// TIA Portal project "Project112" (V16)

(* hardware
DEVICE "S71500/ET200MP station_1"  S7-1500 station
   slot 0: "Rail_0"  Rack  6ES7 590-1***0-0AA0
   slot 0: "PS 25W 24VDC_1"  PS 25W 24VDC  6ES7 505-0KA00-0AB0  V1.0
   slot 1: "fillingStation"  CPU 1511F-1 PN  6ES7 511-1FK00-0AB0  V1.8
      slot 3: "CPU display_1"  6ES7591-1AA00-0AA0
      slot 32768: "PROFINET interface_1"  X1
         slot 32769: "Port_1"  X1 P1
         slot 32770: "Port_2"  X1 P2
   slot 2: "DI 16x24VDC BA_1"  DI 16x24VDC BA  6ES7 521-1BH10-0AA0  V1.1
   slot 3: "DQ 8x24VDC/2A HF_1"  DQ 8x24VDC/2A HF  6ES7 522-1BF00-0AB0  V2.2
   slot 4: "AI 4xU/I/RTD/TC ST_1"  AI 4xU/I/RTD/TC ST  6ES7 531-7QD00-0AB0  V1.0
DEVICE "HMI_1"  TP700 Comfort
   slot 0: "HMI_1"  TP700 Comfort  6AV2 124-0GC01-0AX0  16.0.0.0
   slot 1: "HMI_RT_1"  TP700 Comfort  6AV2 124-0GC01-0AX0  16.0.0.0
   slot 5: "HMI_1.IE_CP_1"  PROFINET Interface  16.0.0.0
      slot 1: "PROFINET Interface_1"  PROFINET Interface
         slot 1: "Port_1"  Port
         slot 2: "Port_2"  Port
   slot 7: "HMI_1.MPI/DP_CP_1"  MPI/DP Interface  16.0.0.0
DEVICE "GSD device_1"  GSD.Device.PN
   slot 0: "Rack"  Rack  V1.0
   slot 0: "SINAMICS-G120-CU240E-2PN"  SINAMICS G120 CU240E-2 PN(-F) V4.5  6SL3 244-0BB1x-1FAx  V4.5
      slot 0: "SINAMICS G120 CU240E-2 PN(-F) V4.5"  SINAMICS G120 CU240E-2 PN(-F) V4.5
      slot 1: "PN-IO"  PN-IO
         slot 1: "Port 1"  Port 1
         slot 2: "Port 2"  Port 2
      slot 1: "Drive_1"  Drive
         slot 0: "Module Access Point"  Module Access Point
   slot 2: "Free telegram, PZD-8/8"  Free telegram, PZD-8/8
*)

// ===== PLC "fillingStation"  CPU 1511F-1 PN =====

VAR_GLOBAL   // PLC tag table "Default tag table"
   "Emg_stop" AT %I0.0 : Bool;
   "Start" AT %I0.1 : Bool;
   "b01_highlevel" AT %I0.2 : Bool;
   "bo2_lowlevel" AT %I0.3 : Bool;
   "pompe_km1" AT %Q0.0 : Bool;
   "valvefilling_1" AT %Q0.1 : Bool;
   "valvefilling_2" AT %Q0.2 : Bool;
   "evacuation_valve" AT %Q0.3 : Bool;
   "stop_bt" AT %M0.0 : Bool;
   "stop_bt(1)" AT %M0.7 : Bool;
   "statehandler" AT %M0.1 : Bool;
   "generalErrors" AT %MD10 : DWord;
   "pompeerror" AT %M10.0 : Bool;
   "pompe_error" AT %M0.2 : Bool;
   "System_Byte" AT %MB1 : Byte;
   "FirstScan" AT %M1.0 : Bool;
   "DiagStatusUpdate" AT %M1.1 : Bool;
   "AlwaysTRUE" AT %M1.2 : Bool;
   "AlwaysFALSE" AT %M1.3 : Bool;
   "System_Byte(1)" AT %MB1 : Byte;
   "Clock_Byte" AT %MB0 : Byte;
   "Clock_10Hz" AT %M0.0 : Bool;
   "Clock_5Hz" AT %M0.1 : Bool;
   "Clock_2.5Hz" AT %M0.2 : Bool;
   "Clock_2Hz" AT %M0.3 : Bool;
   "Clock_1.25Hz" AT %M0.4 : Bool;
   "Clock_1Hz" AT %M0.5 : Bool;
   "Clock_0.625Hz" AT %M0.6 : Bool;
   "Clock_0.5Hz" AT %M0.7 : Bool;
   "actual_wight_card" AT %IW2 : Int;
END_VAR

VAR_GLOBAL   // PLC tag table "input"
   "start(1)" AT %I0.4 : Bool;
   "stop" AT %I0.5 : Bool;
   "reset" AT %I0.6 : Bool;
   "box_detection" AT %I0.7 : Bool;
   "box_at_filling" AT %I1.0 : Bool;
   "box_at_scale" AT %I1.1 : Bool;
   "box_reject" AT %I1.2 : Bool;
   "box_left" AT %I1.3 : Bool;
   "reject_cyl_extended" AT %I1.4 : Bool;
   "reject_cyl_retracted" AT %I1.5 : Bool;
   "caping_cylinder_extended" AT %I1.6 : Bool;
   "caping_cylinder_retracted" AT %I1.7 : Bool;
   "inspect_ol" AT %I2.0 : Bool;
   "conveyer_moving" AT %I2.1 : Bool;
   "valve_switch_open" AT %I2.2 : Bool;
   "main_air_switch" AT %I2.7 : Bool;
   "main_valve_open_fb" AT %I3.1 : Bool;
   "input_vfd" AT %I500.0 : "udt_vfd_status";
   "filling_cyl_retracted" AT %I4.0 : Bool;
   "filling_cyl_extended" AT %I4.1 : Bool;
   "curent_speed" AT %IW600 : Word;
   "part_at_sealing" AT %I3.2 : Bool;
   "cap_carrier_extended" AT %I4.2 : Bool;
   "cap_carrier_retracted" AT %I4.3 : Bool;
   "filling_valve_extended" AT %I4.4 : Bool;
   "filling_valve_retracted" AT %I4.5 : Bool;
   "sealing_locater_extended" AT %I4.6 : Bool;
   "sealing_locater_retacted" AT %I4.7 : Bool;
   "cap_valve_open" AT %I5.0 : Bool;
   "box_at_reject" AT %I5.1 : Bool;
END_VAR

VAR_GLOBAL   // PLC tag table "output"
   "Ev_valve_refill" AT %Q1.0 : Bool;
   "EV_capping" AT %Q1.1 : Bool;
   "EV_capping_return" AT %Q1.2 : Bool;
   "Ev_reject_cylinder" AT %Q1.3 : Bool;
   "main_air_valve" AT %Q1.4 : Bool;
   "tower_green" AT %Q1.5 : Bool;
   "tower_red" AT %Q1.6 : Bool;
   "tower_orange" AT %Q1.7 : Bool;
   "tower_buzer" AT %Q2.0 : Bool;
   "udt_vfd_cmd" AT %Q500.0 : "vfd_cmd";
   "ev_filling_cylinder" AT %Q2.1 : Bool;
   "set_point_vfd" AT %QW600 : Word;
   "cap_motor" AT %Q2.2 : Bool;
   "ev_filling_valve_cyl" AT %Q2.3 : Bool;
   "ev_cap_valve_carrier_cyl" AT %Q2.4 : Bool;
END_VAR

TYPE "udt_state_handler"
   STRUCT
      status : Struct
         ready : Bool;
         running : Bool;
         faulted : Bool;
         stop : Bool;
         safety_ok : Bool;
         air_ok : Bool;
      END_STRUCT;
      cmd : Struct
         reset : Bool;
         start : Bool;
         stop : Bool;
      END_STRUCT;
      cnf : Struct
         state : Int;
      END_STRUCT;
      flts : Struct
         air_system_faulted : Bool;
         safety_emg_stop_btn : Bool;
      END_STRUCT;
   END_STRUCT;
END_TYPE

TYPE "udt_tower_handler"
   STRUCT
      status : Struct
         running : Bool;
         faulted : Bool;
         stop : Bool;
      END_STRUCT;
      cmd : Struct
         turn_red : Bool;
         turn_green : Bool;
         turn_orange : Bool;
         turn_bazer : Bool;
      END_STRUCT;
      flt : Struct
         x_sparte : Bool;
      END_STRUCT;
      cnf : Struct
         x_spare : Bool;
      END_STRUCT;
   END_STRUCT;
END_TYPE

TYPE "udt_equipement"
   STRUCT
      state : Struct
         running : Bool;
         reject_done : Bool;
         filling_done : Bool;
         sealing_done : Bool;
         varification_done : Bool;
         faulted : Bool;
         ready : Bool;
         part_detected : Bool;
         state : Int;
      END_STRUCT;
      cmd : Struct
         converyer_cmd : Bool;
         "filling _valve_cmd" : Bool;
         cmd_cylinder_filling : Bool;
         cmd_cylinder_sealing : Bool;
         cmd_sealing_motor : Bool;
         cmd_cylinder_reject : Bool;
         cmd_trigger_verificaiton : Bool;
         enable_filling : Bool;
         enable_sealing : Bool;
         enable_verification : Bool;
         enable_reject : Bool;
      END_STRUCT;
      flt : Struct
         main_sequece_timeout : Bool;
      END_STRUCT;
      cnf : Struct
         scale_pass_weight : Int := 200;
      END_STRUCT;
   END_STRUCT;
END_TYPE

TYPE "filling_station_udt"
   STRUCT
      status : Struct
         cyl_at_retract : Bool;
         cyl_at_extened : Bool;
         part_at_felling : Bool;
         running : Bool;
         faulted : Bool;
         felling_done : Bool;
         felling_start : Bool;
         valve_open : Bool;
         cyl_valve_at_retract : Bool;
         cyl_valve_at_extend : Bool;
         state : Int;
      END_STRUCT;
      cmd : Struct
         locater_cylinder_cmd : Bool;
         valve_open_cmd : Bool;
         valve_cylinder_cmd : Bool;
      END_STRUCT;
      flt_valve : Word;   // these will define the faults of the valve
      flt2 : Word;   // these are for the filling valve carrier cylinder
      flt1 : Word;   // these are for filling locater cylinder
      cfg : Struct
         valve_open_time : Time := T#10ms;
      END_STRUCT;
   END_STRUCT;
END_TYPE

TYPE "sealing_udt"
   STRUCT
      status : Struct
         cap_carrier_retract : Bool;
         cap_carrier_extended : Bool;
         cyl_at_retract : Bool;
         cyl_at_extended : Bool;
         running : Bool;
         stoped : Bool;
         part_at_sealing : Bool;
         motor_running : Bool;
         cap_present : Bool;
         state : Int;
         open_cap_valve : Int;
      END_STRUCT;
      cmd : Struct
         motor_start_cmd : Bool;
         locater_cyl_cmd : Bool;
         cap_carring_cyl_cmd : Bool;
         open_cap_valve_cmd : Bool;
      END_STRUCT;
      flt_valve : Word;
      flt_valve_carrier_cyl : Word;
      flt_locater_cylinder : Word;
      cnf : Struct
         spare : Bool;
      END_STRUCT;
   END_STRUCT;
END_TYPE

TYPE "scaling_udt"
   STRUCT
      status : Struct
         actual_weight_bottle : Int;
         running : Bool;
         stop : Bool;
         pass_part : Bool;
         reject_part : Bool;
      END_STRUCT;
      cmd : Struct
         spare : Bool;
      END_STRUCT;
      cnf : Struct
         max_weight : Int := 140;
         min_weight : Int := 150;
      END_STRUCT;
      flt : Word;
   END_STRUCT;
END_TYPE

TYPE "reject_udt"
   STRUCT
      status : Struct
         cyl_at_retract : Bool;
         cyl_at_extend : Bool;
         running : Bool;
         faulted : Bool;
         state : Int;
      END_STRUCT;
      cmd : Struct
         spare : Bool;
      END_STRUCT;
      flt : Word;
      cnf : Struct
         reject_count : Int;
      END_STRUCT;
   END_STRUCT;
END_TYPE

TYPE "udt_vfd_status"
   STRUCT
      "Ready to switch on" : Bool;
      "Ready for operation" : Bool;
      "Operation enabled" : Bool;
      "Fault active" : Bool;
      "OFF2 inactive" : Bool;
      "OFF3 inactive" : Bool;
      "Switching-on inhibited" : Bool;
      "Warning active" : Bool;
      "Speed setpoint/actual value comparison" : Bool;
      "Control requested" : Bool;
      "Setpoint reached" : Bool;
      "Torque limit active" : Bool;
   END_STRUCT;
END_TYPE

TYPE "vfd_cmd"
   STRUCT
      "ON/OFF1" : Bool;
      OFF2 : Bool;
      OFF3 : Bool;
      "Enable operation" : Bool;
      "Enable ramp-function generator" : Bool;
      "Continue ramp-function generator" : Bool;
      "Enable setpoint" : Bool;
      "Acknowledge fault" : Bool;
      "Control by PLC" : Bool;
   END_STRUCT;
END_TYPE

TYPE "hmi_cmd_state"
   STRUCT
      cmd : Struct
         oprator_speed_setpoint : Int;
      END_STRUCT;
      status : Struct
         set_point_valid : Bool;
      END_STRUCT;
   END_STRUCT;
END_TYPE

DATA_BLOCK "Main_Safety_RTG1_DB"   // DB1, F_DB
{ S7_Optimized_Access := 'TRUE' }
NAME : FUSI
VERSION : 0.1
// stored: InstanceOfName Main_Safety_RTG1
"Main_Safety_RTG1"
BEGIN
END_DATA_BLOCK

DATA_BLOCK "global_data_block"   // DB6
{ S7_Optimized_Access := 'TRUE' }
VERSION : 0.1
   VAR
      verification_handler : "scaling_udt";
      reject_handler : "reject_udt";
      hmi_cmd_state : "hmi_cmd_state";
      sealing_handler : "sealing_udt";
      equipement_handler : "udt_equipement";
      filling_station_handler : "filling_station_udt";
      tower_handling : "udt_tower_handler";
      machine_state : "udt_state_handler";
   END_VAR
BEGIN
END_DATA_BLOCK

// folder: System blocks/Program resources

DATA_BLOCK "air_check"   // DB2
{ S7_Optimized_Access := 'TRUE' }
AUTHOR : Simatic
FAMILY : IEC
NAME : IEC_TMR
VERSION : 1.0
// stored: InstanceOfName IEC_TIMER
"IEC_TIMER"
BEGIN
END_DATA_BLOCK

DATA_BLOCK "verify_air_present"   // DB5
{ S7_Optimized_Access := 'TRUE' }
AUTHOR : Simatic
FAMILY : IEC
NAME : IEC_TMR
VERSION : 1.0
// stored: InstanceOfName IEC_TIMER
"IEC_TIMER"
BEGIN
END_DATA_BLOCK

DATA_BLOCK "valve_timing"   // DB15
{ S7_Optimized_Access := 'TRUE' }
AUTHOR : Simatic
FAMILY : IEC
NAME : IEC_TMR
VERSION : 1.0
// stored: InstanceOfName IEC_TIMER
"IEC_TIMER"
BEGIN
END_DATA_BLOCK

DATA_BLOCK "IEC_Timer_0_DB_1"   // DB16
{ S7_Optimized_Access := 'TRUE' }
AUTHOR : Simatic
FAMILY : IEC
NAME : IEC_TMR
VERSION : 1.0
// stored: InstanceOfName IEC_TIMER
"IEC_TIMER"
BEGIN
END_DATA_BLOCK

DATA_BLOCK "motor_time"   // DB17
{ S7_Optimized_Access := 'TRUE' }
AUTHOR : Simatic
FAMILY : IEC
NAME : IEC_TMR
VERSION : 1.0
// stored: InstanceOfName IEC_TIMER
"IEC_TIMER"
BEGIN
END_DATA_BLOCK

DATA_BLOCK "IEC_Timer_0_DB_2"   // DB18
{ S7_Optimized_Access := 'TRUE' }
AUTHOR : Simatic
FAMILY : IEC
NAME : IEC_TMR
VERSION : 1.0
// stored: InstanceOfName IEC_TIMER
"IEC_TIMER"
BEGIN
END_DATA_BLOCK

DATA_BLOCK "IEC_Timer_0_DB_3"   // DB19
{ S7_Optimized_Access := 'TRUE' }
AUTHOR : Simatic
FAMILY : IEC
NAME : IEC_TMR
VERSION : 1.0
// stored: InstanceOfName IEC_TIMER
"IEC_TIMER"
BEGIN
END_DATA_BLOCK

DATA_BLOCK "wire_break"   // DB20
{ S7_Optimized_Access := 'TRUE' }
AUTHOR : Simatic
FAMILY : IEC
NAME : IEC_TMR
VERSION : 1.0
// stored: InstanceOfName IEC_TIMER
"IEC_TIMER"
BEGIN
END_DATA_BLOCK

DATA_BLOCK "IEC_Timer_0_DB_4"   // DB21
{ S7_Optimized_Access := 'TRUE' }
AUTHOR : Simatic
FAMILY : IEC
NAME : IEC_TMR
VERSION : 1.0
// stored: InstanceOfName IEC_TIMER
"IEC_TIMER"
BEGIN
END_DATA_BLOCK

DATA_BLOCK "IEC_Timer_0_DB_5"   // DB22
{ S7_Optimized_Access := 'TRUE' }
AUTHOR : Simatic
FAMILY : IEC
NAME : IEC_TMR
VERSION : 1.0
// stored: InstanceOfName IEC_TIMER
"IEC_TIMER"
BEGIN
END_DATA_BLOCK

DATA_BLOCK "timeout]"   // DB25
{ S7_Optimized_Access := 'TRUE' }
AUTHOR : Simatic
FAMILY : IEC
NAME : IEC_TMR
VERSION : 1.0
// stored: InstanceOfName IEC_TIMER
"IEC_TIMER"
BEGIN
END_DATA_BLOCK

DATA_BLOCK "IEC_Timer_0_DB_8"   // DB26
{ S7_Optimized_Access := 'TRUE' }
AUTHOR : Simatic
FAMILY : IEC
NAME : IEC_TMR
VERSION : 1.0
// stored: InstanceOfName IEC_TIMER
"IEC_TIMER"
BEGIN
END_DATA_BLOCK

DATA_BLOCK "signal_che k"   // DB27
{ S7_Optimized_Access := 'TRUE' }
AUTHOR : Simatic
FAMILY : IEC
NAME : IEC_TMR
VERSION : 1.0
// stored: InstanceOfName IEC_TIMER
"IEC_TIMER"
BEGIN
END_DATA_BLOCK

DATA_BLOCK "cyl_extended_check"   // DB28
{ S7_Optimized_Access := 'TRUE' }
AUTHOR : Simatic
FAMILY : IEC
NAME : IEC_TMR
VERSION : 1.0
// stored: InstanceOfName IEC_TIMER
"IEC_TIMER"
BEGIN
END_DATA_BLOCK

DATA_BLOCK "cylinder"   // DB29
{ S7_Optimized_Access := 'TRUE' }
AUTHOR : Simatic
FAMILY : IEC
NAME : IEC_TMR
VERSION : 1.0
// stored: InstanceOfName IEC_TIMER
"IEC_TIMER"
BEGIN
END_DATA_BLOCK

DATA_BLOCK "IEC_Timer_0_DB_9"   // DB30
{ S7_Optimized_Access := 'TRUE' }
AUTHOR : Simatic
FAMILY : IEC
NAME : IEC_TMR
VERSION : 1.0
// stored: InstanceOfName IEC_TIMER
"IEC_TIMER"
BEGIN
END_DATA_BLOCK

DATA_BLOCK "setpoint"   // DB31
{ S7_Optimized_Access := 'TRUE' }
AUTHOR : Simatic
FAMILY : IEC
NAME : IEC_TMR
VERSION : 1.0
// stored: InstanceOfName IEC_TIMER
"IEC_TIMER"
BEGIN
END_DATA_BLOCK

DATA_BLOCK "IEC_Timer_0_DB_10"   // DB33
{ S7_Optimized_Access := 'TRUE' }
AUTHOR : Simatic
FAMILY : IEC
NAME : IEC_TMR
VERSION : 1.0
// stored: InstanceOfName IEC_TIMER
"IEC_TIMER"
BEGIN
END_DATA_BLOCK

// folder: equipement

DATA_BLOCK "filling_sequence_DB"   // DB11
{ S7_Optimized_Access := 'TRUE' }
VERSION : 0.1
// stored: InstanceOfName filling_sequence
"filling_sequence"
BEGIN
END_DATA_BLOCK

DATA_BLOCK "sealing_db"   // DB12
{ S7_Optimized_Access := 'TRUE' }
VERSION : 0.1
// stored: InstanceOfName sealing_sequnce
"sealing_sequnce"
BEGIN
END_DATA_BLOCK

DATA_BLOCK "scaling_sequence_DB"   // DB13
{ S7_Optimized_Access := 'TRUE' }
VERSION : 0.1
// stored: InstanceOfName scaling_sequence
"scaling_sequence"
BEGIN
END_DATA_BLOCK

DATA_BLOCK "1_main_squence_DB"   // DB32
{ S7_Optimized_Access := 'TRUE' }
VERSION : 0.1
// stored: InstanceOfName 1_main_squence
"1_main_squence"
BEGIN
END_DATA_BLOCK

// folder: machine

DATA_BLOCK "safety_block_DB"   // DB7
{ S7_Optimized_Access := 'TRUE' }
VERSION : 0.1
// stored: InstanceOfName safety_block
"safety_block"
BEGIN
END_DATA_BLOCK

DATA_BLOCK "air_management_blk_DB"   // DB8
{ S7_Optimized_Access := 'TRUE' }
VERSION : 0.1
// stored: InstanceOfName air_management_blk
"air_management_blk"
BEGIN
END_DATA_BLOCK

DATA_BLOCK "tower_handler_DB"   // DB9
{ S7_Optimized_Access := 'TRUE' }
VERSION : 0.1
// stored: InstanceOfName tower_handler
"tower_handler"
BEGIN
END_DATA_BLOCK

DATA_BLOCK "state_handler_DB"   // DB10
{ S7_Optimized_Access := 'TRUE' }
VERSION : 0.1
// stored: InstanceOfName state_handler
"state_handler"
BEGIN
END_DATA_BLOCK

// folder: (top level)

FUNCTION_BLOCK "Main_Safety_RTG1"   // FB1, F_FBD
{ S7_Optimized_Access := 'TRUE' }
BEGIN

REGION Network 1
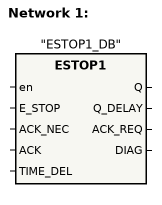
   "ESTOP1_DB"();   // ESTOP1
END_REGION
END_FUNCTION_BLOCK

ORGANIZATION_BLOCK "Main"   // OB1, LAD, ProgramCycle
TITLE = "Main Program Sweep (Cycle)"
{ S7_Optimized_Access := 'TRUE' }
VERSION : 0.1
   VAR_INPUT
      Initial_Call : Bool;   // Initial call of this OB
      Remanence : Bool;   // =True, if remanent data are available
   END_VAR
BEGIN

REGION Network 1: this the systeme process
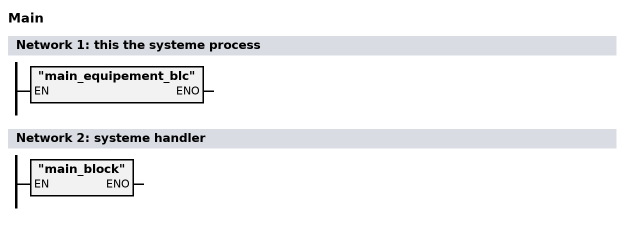
   RUNG wire#powerrail
      "main_equipement_blc"()
   END_RUNG
   // the same network as SCL:
   "main_equipement_blc"();
END_REGION

REGION Network 2: systeme handler
   RUNG wire#powerrail
      "main_block"()
   END_RUNG
   // the same network as SCL:
   "main_block"();
END_REGION

REGION Network 3: error handler block
END_REGION
END_ORGANIZATION_BLOCK

// folder: equipement

FUNCTION_BLOCK "1_main_squence"   // FB6, LAD
{ S7_Optimized_Access := 'TRUE' }
VERSION : 0.1
   VAR_INPUT
      conveyor_feedbak : Bool;
      part_at_filling : Bool;
      part_at_sealing : Bool;
      part_verification : Bool;
      part_at_reject : Bool;
   END_VAR
   VAR_IN_OUT
      equipement_handler : "udt_equipement";
      machine_handler : "udt_state_handler";
   END_VAR
   VAR
      cycle_lock : Bool;
      bottle_count_done : Int;
      reject_instance : "reject_main";
   END_VAR
   VAR_TEMP
      bottle_done_process : Bool;
      bottle_succesed : Bool;
   END_VAR
   VAR_TEMP   // added for the SCL form of the ladder/FBD networks
      _w1 : Bool;
      _w2 : Bool;
      _w3 : Bool;
      _w4 : Bool;
      _w5 : Bool;
      _w6 : Bool;
      _w7 : Bool;
   END_VAR
BEGIN

REGION Network 1: move the machine from idle to running state
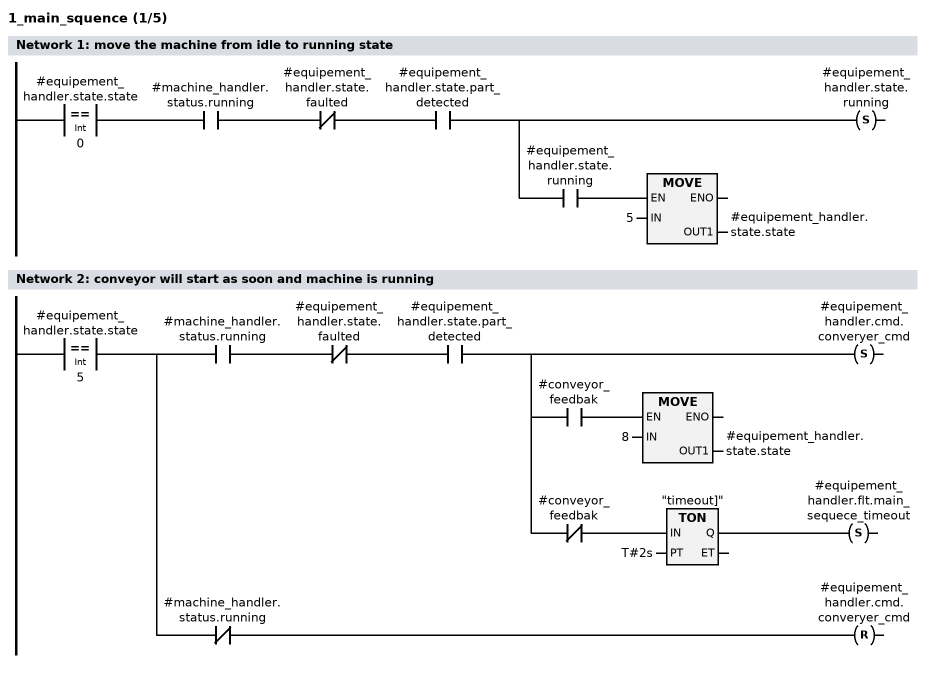
   RUNG wire#powerrail
      { S7_Templates := "SrcType := Int" } EQ_Contact(in1 := #equipement_handler.state.state, in2 := 0)
      Contact( #machine_handler.status.running )
      I_Contact( #equipement_handler.state.faulted )
      Contact( #equipement_handler.state.part_detected )
      wire#w1
      S_Coil( #equipement_handler.state.running )
   END_RUNG
   RUNG wire#w1
      Contact( #equipement_handler.state.running )
      Move(in := 5, out1 => #equipement_handler.state.state)
   END_RUNG
   // the same network as SCL:
   #_w1 := (#equipement_handler.state.state = 0) AND #machine_handler.status.running AND NOT #equipement_handler.state.faulted AND #equipement_handler.state.part_detected;
   IF #_w1 THEN #equipement_handler.state.running := TRUE; END_IF;
   IF #_w1 AND #equipement_handler.state.running THEN #equipement_handler.state.state := 5; END_IF;
END_REGION

REGION Network 2: conveyor will start as soon and machine is running
   #_w1 := #equipement_handler.state.state = 5;
   #_w2 := #_w1 AND #machine_handler.status.running AND NOT #equipement_handler.state.faulted AND #equipement_handler.state.part_detected;
   IF #_w2 THEN #equipement_handler.cmd.converyer_cmd := TRUE; END_IF;
   IF #_w2 AND #conveyor_feedbak THEN #equipement_handler.state.state := 8; END_IF;
   "timeout]".TON(IN := #_w2 AND NOT #conveyor_feedbak, PT := T#2s);
   IF "timeout]".Q THEN #equipement_handler.flt.main_sequece_timeout := TRUE; END_IF;
   IF #_w1 AND NOT #machine_handler.status.running THEN
       #equipement_handler.cmd.converyer_cmd := FALSE;
   END_IF;
END_REGION

REGION Network 3: 5 according which sensor gets triggered different station will be enabled
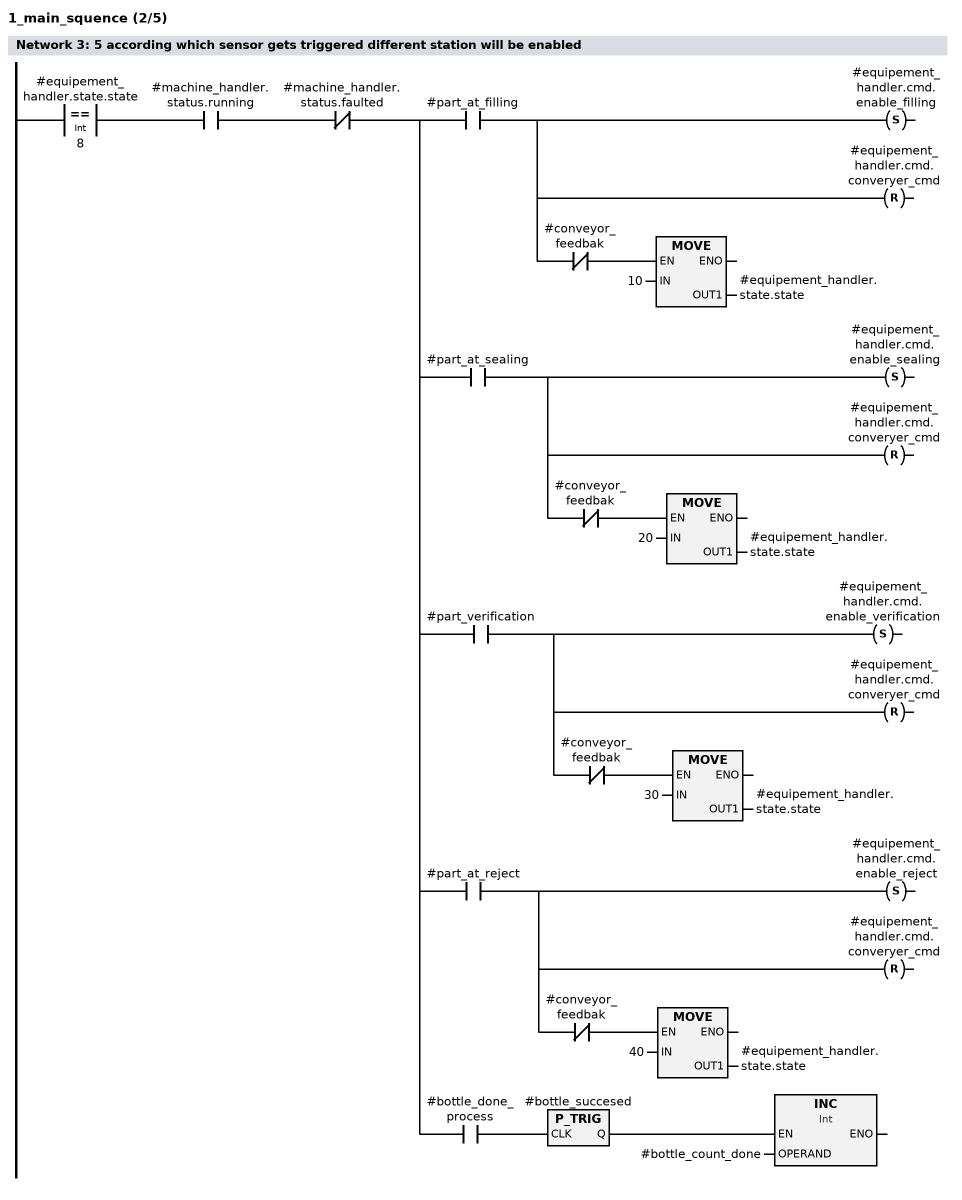
   RUNG wire#powerrail
      { S7_Templates := "SrcType := Int" } EQ_Contact(in1 := #equipement_handler.state.state, in2 := 8)
      Contact( #machine_handler.status.running )
      I_Contact( #machine_handler.status.faulted )
      wire#w1
      Contact( #part_at_filling )
      wire#w2
      S_Coil( #equipement_handler.cmd.enable_filling )
   END_RUNG
   RUNG wire#w2
      R_Coil( #equipement_handler.cmd.converyer_cmd )
   END_RUNG
   RUNG wire#w2
      I_Contact( #conveyor_feedbak )
      Move(in := 10, out1 => #equipement_handler.state.state)
   END_RUNG
   RUNG wire#w1
      Contact( #part_at_sealing )
      wire#w3
      S_Coil( #equipement_handler.cmd.enable_sealing )
   END_RUNG
   RUNG wire#w3
      R_Coil( #equipement_handler.cmd.converyer_cmd )
   END_RUNG
   RUNG wire#w3
      I_Contact( #conveyor_feedbak )
      Move(in := 20, out1 => #equipement_handler.state.state)
   END_RUNG
   RUNG wire#w1
      Contact( #part_verification )
      wire#w4
      S_Coil( #equipement_handler.cmd.enable_verification )
   END_RUNG
   RUNG wire#w4
      R_Coil( #equipement_handler.cmd.converyer_cmd )
   END_RUNG
   RUNG wire#w4
      I_Contact( #conveyor_feedbak )
      Move(in := 30, out1 => #equipement_handler.state.state)
   END_RUNG
   RUNG wire#w1
      Contact( #part_at_reject )
      wire#w5
      S_Coil( #equipement_handler.cmd.enable_reject )
   END_RUNG
   RUNG wire#w5
      R_Coil( #equipement_handler.cmd.converyer_cmd )
   END_RUNG
   RUNG wire#w5
      I_Contact( #conveyor_feedbak )
      Move(in := 40, out1 => #equipement_handler.state.state)
   END_RUNG
   RUNG wire#w1
      Contact( #bottle_done_process )
      P_Trig( #bottle_succesed )
      { S7_Templates := "DestType := Int" } Inc( #bottle_count_done )
   END_RUNG
   // the same network as SCL:
   #_w1 := (#equipement_handler.state.state = 8) AND #machine_handler.status.running AND NOT #machine_handler.status.faulted;
   #_w2 := #_w1 AND #part_at_filling;
   IF #_w2 THEN
       #equipement_handler.cmd.enable_filling := TRUE;
       #equipement_handler.cmd.converyer_cmd := FALSE;
   END_IF;
   IF #_w2 AND NOT #conveyor_feedbak THEN #equipement_handler.state.state := 10; END_IF;
   #_w3 := #_w1 AND #part_at_sealing;
   IF #_w3 THEN
       #equipement_handler.cmd.enable_sealing := TRUE;
       #equipement_handler.cmd.converyer_cmd := FALSE;
   END_IF;
   IF #_w3 AND NOT #conveyor_feedbak THEN #equipement_handler.state.state := 20; END_IF;
   #_w4 := #_w1 AND #part_verification;
   IF #_w4 THEN
       #equipement_handler.cmd.enable_verification := TRUE;
       #equipement_handler.cmd.converyer_cmd := FALSE;
   END_IF;
   IF #_w4 AND NOT #conveyor_feedbak THEN #equipement_handler.state.state := 30; END_IF;
   #_w5 := #_w1 AND #part_at_reject;
   IF #_w5 THEN
       #equipement_handler.cmd.enable_reject := TRUE;
       #equipement_handler.cmd.converyer_cmd := FALSE;
   END_IF;
   IF #_w5 AND NOT #conveyor_feedbak THEN #equipement_handler.state.state := 40; END_IF;
   #_w6 := #_w1 AND #bottle_done_process;
   #_w7 := #_w6 AND NOT #bottle_succesed;   // rising edge
   #bottle_succesed := #_w6;
   IF #_w7 THEN #bottle_count_done := #bottle_count_done + 1; END_IF;
END_REGION

REGION Network 4: 10 call the filling process
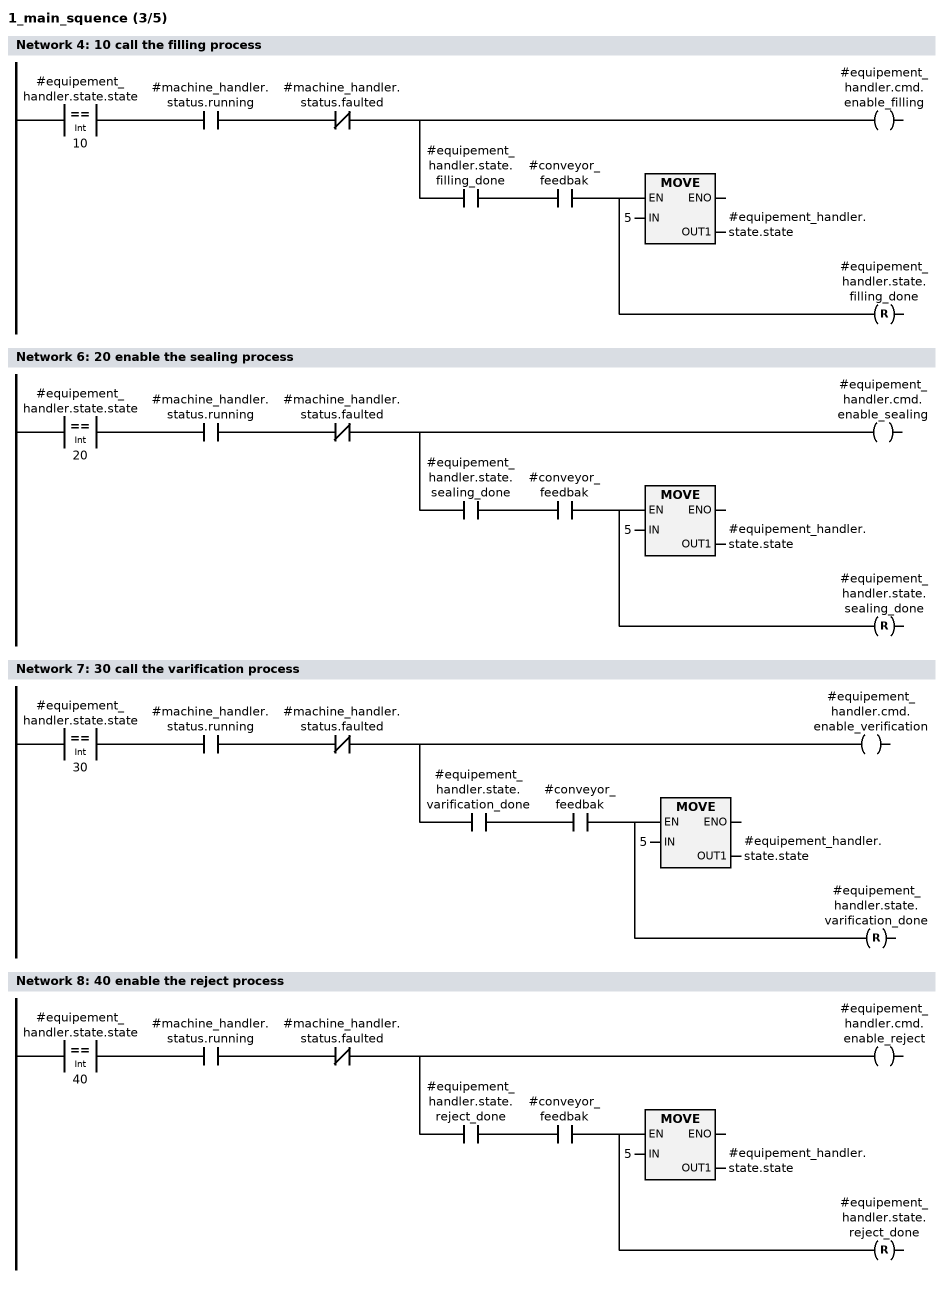
   RUNG wire#powerrail
      { S7_Templates := "SrcType := Int" } EQ_Contact(in1 := #equipement_handler.state.state, in2 := 10)
      Contact( #machine_handler.status.running )
      I_Contact( #machine_handler.status.faulted )
      wire#w1
      Coil( #equipement_handler.cmd.enable_filling )
   END_RUNG
   RUNG wire#w1
      Contact( #equipement_handler.state.filling_done )
      Contact( #conveyor_feedbak )
      wire#w2
      Move(in := 5, out1 => #equipement_handler.state.state)
   END_RUNG
   RUNG wire#w2
      R_Coil( #equipement_handler.state.filling_done )
   END_RUNG
   // the same network as SCL:
   #equipement_handler.cmd.enable_filling := (#equipement_handler.state.state = 10) AND #machine_handler.status.running AND NOT #machine_handler.status.faulted;
   IF #equipement_handler.cmd.enable_filling AND #equipement_handler.state.filling_done AND #conveyor_feedbak THEN
       #equipement_handler.state.state := 5;
       #equipement_handler.state.filling_done := FALSE;
   END_IF;
END_REGION

REGION Network 6: 20 enable the sealing process
   RUNG wire#powerrail
      { S7_Templates := "SrcType := Int" } EQ_Contact(in1 := #equipement_handler.state.state, in2 := 20)
      Contact( #machine_handler.status.running )
      I_Contact( #machine_handler.status.faulted )
      wire#w1
      Coil( #equipement_handler.cmd.enable_sealing )
   END_RUNG
   RUNG wire#w1
      Contact( #equipement_handler.state.sealing_done )
      Contact( #conveyor_feedbak )
      wire#w2
      Move(in := 5, out1 => #equipement_handler.state.state)
   END_RUNG
   RUNG wire#w2
      R_Coil( #equipement_handler.state.sealing_done )
   END_RUNG
   // the same network as SCL:
   #equipement_handler.cmd.enable_sealing := (#equipement_handler.state.state = 20) AND #machine_handler.status.running AND NOT #machine_handler.status.faulted;
   IF #equipement_handler.cmd.enable_sealing AND #equipement_handler.state.sealing_done AND #conveyor_feedbak THEN
       #equipement_handler.state.state := 5;
       #equipement_handler.state.sealing_done := FALSE;
   END_IF;
END_REGION

REGION Network 7: 30 call the varification process
   RUNG wire#powerrail
      { S7_Templates := "SrcType := Int" } EQ_Contact(in1 := #equipement_handler.state.state, in2 := 30)
      Contact( #machine_handler.status.running )
      I_Contact( #machine_handler.status.faulted )
      wire#w1
      Coil( #equipement_handler.cmd.enable_verification )
   END_RUNG
   RUNG wire#w1
      Contact( #equipement_handler.state.varification_done )
      Contact( #conveyor_feedbak )
      wire#w2
      Move(in := 5, out1 => #equipement_handler.state.state)
   END_RUNG
   RUNG wire#w2
      R_Coil( #equipement_handler.state.varification_done )
   END_RUNG
   // the same network as SCL:
   #equipement_handler.cmd.enable_verification := (#equipement_handler.state.state = 30) AND #machine_handler.status.running AND NOT #machine_handler.status.faulted;
   IF #equipement_handler.cmd.enable_verification AND #equipement_handler.state.varification_done AND #conveyor_feedbak THEN
       #equipement_handler.state.state := 5;
       #equipement_handler.state.varification_done := FALSE;
   END_IF;
END_REGION

REGION Network 8: 40 enable the reject process
   RUNG wire#powerrail
      { S7_Templates := "SrcType := Int" } EQ_Contact(in1 := #equipement_handler.state.state, in2 := 40)
      Contact( #machine_handler.status.running )
      I_Contact( #machine_handler.status.faulted )
      wire#w1
      Coil( #equipement_handler.cmd.enable_reject )
   END_RUNG
   RUNG wire#w1
      Contact( #equipement_handler.state.reject_done )
      Contact( #conveyor_feedbak )
      wire#w2
      Move(in := 5, out1 => #equipement_handler.state.state)
   END_RUNG
   RUNG wire#w2
      R_Coil( #equipement_handler.state.reject_done )
   END_RUNG
   // the same network as SCL:
   #equipement_handler.cmd.enable_reject := (#equipement_handler.state.state = 40) AND #machine_handler.status.running AND NOT #machine_handler.status.faulted;
   IF #equipement_handler.cmd.enable_reject AND #equipement_handler.state.reject_done AND #conveyor_feedbak THEN
       #equipement_handler.state.state := 5;
       #equipement_handler.state.reject_done := FALSE;
   END_IF;
END_REGION

REGION Network 9: call the filling process
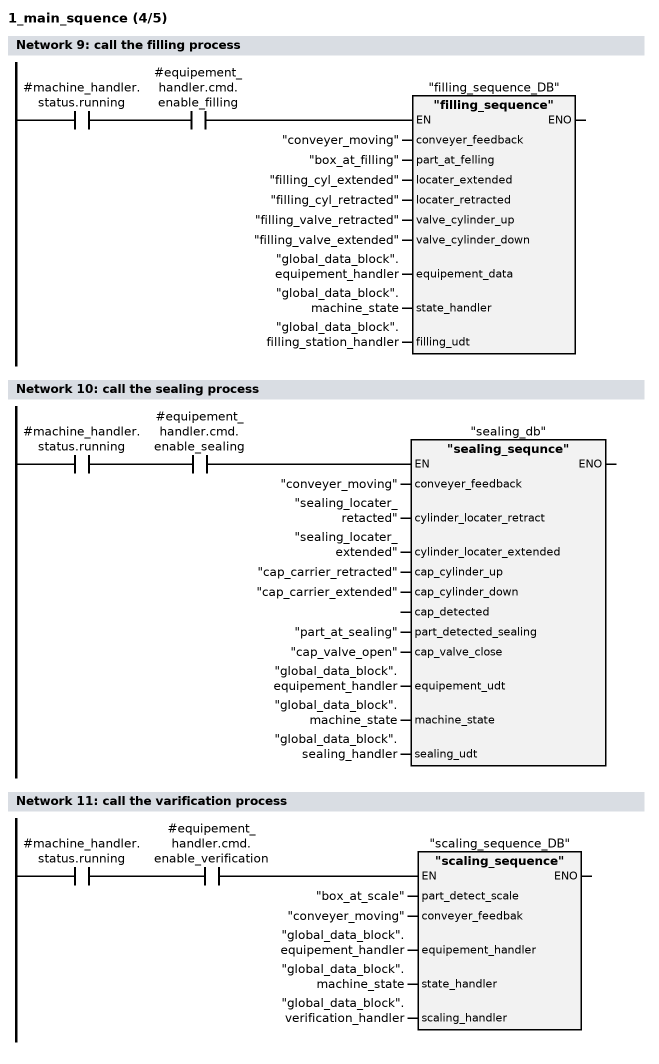
   RUNG wire#powerrail
      Contact( #machine_handler.status.running )
      Contact( #equipement_handler.cmd.enable_filling )
      "filling_sequence_DB"(conveyer_feedback := "conveyer_moving", part_at_felling := "box_at_filling", locater_extended := "filling_cyl_extended", locater_retracted := "filling_cyl_retracted", valve_cylinder_up := "filling_valve_retracted", valve_cylinder_down := "filling_valve_extended", equipement_data := "global_data_block".equipement_handler, state_handler := "global_data_block".machine_state, filling_udt := "global_data_block".filling_station_handler)
   END_RUNG
   // the same network as SCL:
   IF #machine_handler.status.running AND #equipement_handler.cmd.enable_filling THEN
       "filling_sequence_DB"(conveyer_feedback := "conveyer_moving",   // "filling_sequence"
                             part_at_felling := "box_at_filling",
                             locater_extended := "filling_cyl_extended",
                             locater_retracted := "filling_cyl_retracted",
                             valve_cylinder_up := "filling_valve_retracted",
                             valve_cylinder_down := "filling_valve_extended",
                             equipement_data := "global_data_block".equipement_handler,
                             state_handler := "global_data_block".machine_state,
                             filling_udt := "global_data_block".filling_station_handler);
   END_IF;
END_REGION

REGION Network 10: call the sealing process
   RUNG wire#powerrail
      Contact( #machine_handler.status.running )
      Contact( #equipement_handler.cmd.enable_sealing )
      "sealing_db"(conveyer_feedback := "conveyer_moving", cylinder_locater_retract := "sealing_locater_retacted", cylinder_locater_extended := "sealing_locater_extended", cap_cylinder_up := "cap_carrier_retracted", cap_cylinder_down := "cap_carrier_extended", cap_detected :=, part_detected_sealing := "part_at_sealing", cap_valve_close := "cap_valve_open", equipement_udt := "global_data_block".equipement_handler, machine_state := "global_data_block".machine_state, sealing_udt := "global_data_block".sealing_handler)
   END_RUNG
   // the same network as SCL:
   IF #machine_handler.status.running AND #equipement_handler.cmd.enable_sealing THEN
       "sealing_db"(conveyer_feedback := "conveyer_moving",   // "sealing_sequnce"
                    cylinder_locater_retract := "sealing_locater_retacted",
                    cylinder_locater_extended := "sealing_locater_extended",
                    cap_cylinder_up := "cap_carrier_retracted",
                    cap_cylinder_down := "cap_carrier_extended",
                    part_detected_sealing := "part_at_sealing",
                    cap_valve_close := "cap_valve_open",
                    equipement_udt := "global_data_block".equipement_handler,
                    machine_state := "global_data_block".machine_state,
                    sealing_udt := "global_data_block".sealing_handler);
   END_IF;
END_REGION

REGION Network 11: call the varification process
   RUNG wire#powerrail
      Contact( #machine_handler.status.running )
      Contact( #equipement_handler.cmd.enable_verification )
      "scaling_sequence_DB"(part_detect_scale := "box_at_scale", conveyer_feedbak := "conveyer_moving", equipement_handler := "global_data_block".equipement_handler, state_handler := "global_data_block".machine_state, scaling_handler := "global_data_block".verification_handler)
   END_RUNG
   // the same network as SCL:
   IF #machine_handler.status.running AND #equipement_handler.cmd.enable_verification THEN
       "scaling_sequence_DB"(part_detect_scale := "box_at_scale",   // "scaling_sequence"
                             conveyer_feedbak := "conveyer_moving",
                             equipement_handler := "global_data_block".equipement_handler,
                             state_handler := "global_data_block".machine_state,
                             scaling_handler := "global_data_block".verification_handler);
   END_IF;
END_REGION

REGION Network 12: call the reject process
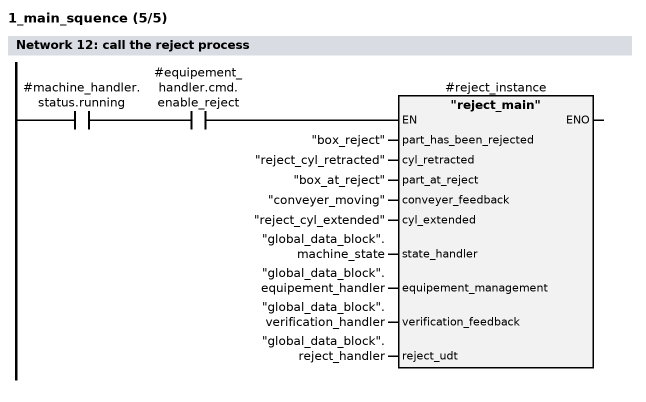
   RUNG wire#powerrail
      Contact( #machine_handler.status.running )
      Contact( #equipement_handler.cmd.enable_reject )
      #reject_instance(part_has_been_rejected := "box_reject", cyl_retracted := "reject_cyl_retracted", part_at_reject := "box_at_reject", conveyer_feedback := "conveyer_moving", cyl_extended := "reject_cyl_extended", state_handler := "global_data_block".machine_state, equipement_management := "global_data_block".equipement_handler, verification_feedback := "global_data_block".verification_handler, reject_udt := "global_data_block".reject_handler)
   END_RUNG
   // the same network as SCL:
   IF #machine_handler.status.running AND #equipement_handler.cmd.enable_reject THEN
       #reject_instance(part_has_been_rejected := "box_reject",   // "reject_main"
                        cyl_retracted := "reject_cyl_retracted",
                        part_at_reject := "box_at_reject",
                        conveyer_feedback := "conveyer_moving",
                        cyl_extended := "reject_cyl_extended",
                        state_handler := "global_data_block".machine_state,
                        equipement_management := "global_data_block".equipement_handler,
                        verification_feedback := "global_data_block".verification_handler,
                        reject_udt := "global_data_block".reject_handler);
   END_IF;
END_REGION
END_FUNCTION_BLOCK

FUNCTION "main_equipement_blc" : Void   // FC2, LAD
{ S7_Optimized_Access := 'TRUE' }
VERSION : 0.1
BEGIN

REGION Network 1: call the main process control block
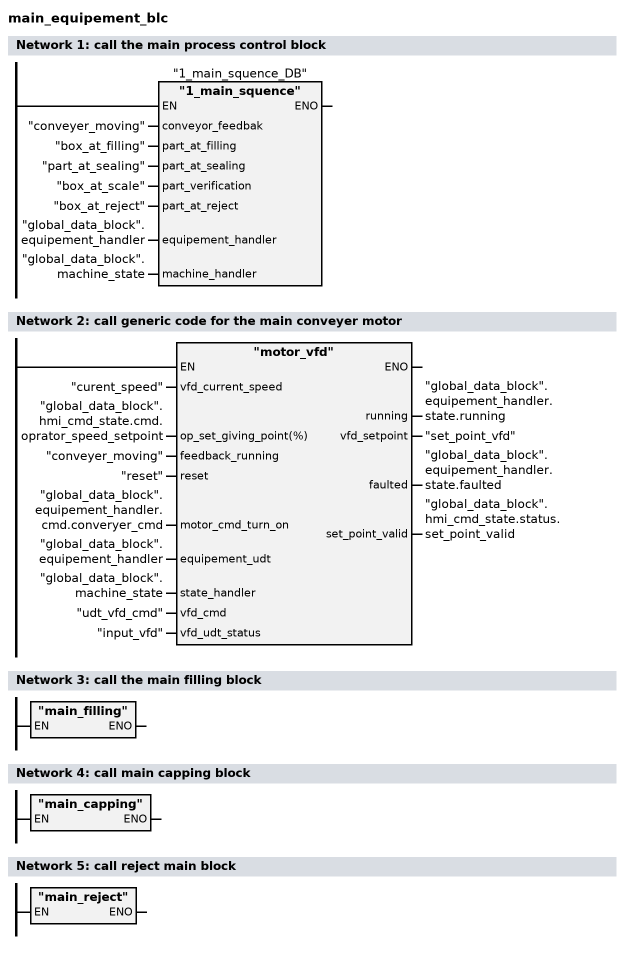
   RUNG wire#powerrail
      "1_main_squence_DB"(conveyor_feedbak := "conveyer_moving", part_at_filling := "box_at_filling", part_at_sealing := "part_at_sealing", part_verification := "box_at_scale", part_at_reject := "box_at_reject", equipement_handler := "global_data_block".equipement_handler, machine_handler := "global_data_block".machine_state)
   END_RUNG
   // the same network as SCL:
   "1_main_squence_DB"(conveyor_feedbak := "conveyer_moving",   // "1_main_squence"
                       part_at_filling := "box_at_filling",
                       part_at_sealing := "part_at_sealing",
                       part_verification := "box_at_scale",
                       part_at_reject := "box_at_reject",
                       equipement_handler := "global_data_block".equipement_handler,
                       machine_handler := "global_data_block".machine_state);
END_REGION

REGION Network 2: call generic code for the main conveyer motor
   RUNG wire#powerrail
      "motor_vfd"(vfd_current_speed := "curent_speed", "op_set_giving_point(%)" := "global_data_block".hmi_cmd_state.cmd.oprator_speed_setpoint, feedback_running := "conveyer_moving", reset := "reset", motor_cmd_turn_on := "global_data_block".equipement_handler.cmd.converyer_cmd, equipement_udt := "global_data_block".equipement_handler, state_handler := "global_data_block".machine_state, vfd_cmd := "udt_vfd_cmd", vfd_udt_status := "input_vfd", running => "global_data_block".equipement_handler.state.running, vfd_setpoint => "set_point_vfd", faulted => "global_data_block".equipement_handler.state.faulted, set_point_valid => "global_data_block".hmi_cmd_state.status.set_point_valid)
   END_RUNG
   // the same network as SCL:
   "motor_vfd"(vfd_current_speed := "curent_speed",
               "op_set_giving_point(%)" := "global_data_block".hmi_cmd_state.cmd.oprator_speed_setpoint,
               feedback_running := "conveyer_moving",
               reset := "reset",
               motor_cmd_turn_on := "global_data_block".equipement_handler.cmd.converyer_cmd,
               equipement_udt := "global_data_block".equipement_handler,
               state_handler := "global_data_block".machine_state,
               vfd_cmd := "udt_vfd_cmd",
               vfd_udt_status := "input_vfd",
               running => "global_data_block".equipement_handler.state.running,
               vfd_setpoint => "set_point_vfd",
               faulted => "global_data_block".equipement_handler.state.faulted,
               set_point_valid => "global_data_block".hmi_cmd_state.status.set_point_valid);
END_REGION

REGION Network 3: call the main filling block
   RUNG wire#powerrail
      "main_filling"()
   END_RUNG
   // the same network as SCL:
   "main_filling"();
END_REGION

REGION Network 4: call main capping block
   RUNG wire#powerrail
      "main_capping"()
   END_RUNG
   // the same network as SCL:
   "main_capping"();
END_REGION

REGION Network 5: call reject main block
   RUNG wire#powerrail
      "main_reject"()
   END_RUNG
   // the same network as SCL:
   "main_reject"();
END_REGION
END_FUNCTION

// folder: equipement/capping

FUNCTION_BLOCK "sealing_sequnce"   // FB9, LAD
{ S7_Optimized_Access := 'TRUE' }
VERSION : 0.1
   VAR_INPUT
      conveyer_feedback : Bool;
      cylinder_locater_retract : Bool;
      cylinder_locater_extended : Bool;
      cap_cylinder_up : Bool;
      cap_cylinder_down : Bool;
      cap_detected : Bool;
      part_detected_sealing : Bool;
      cap_valve_close : Bool;
   END_VAR
   VAR_IN_OUT
      equipement_udt : "udt_equipement";
      machine_state : "udt_state_handler";
      sealing_udt : "sealing_udt";
   END_VAR
   VAR
      motor_time_seal : TON_TIME;
      start_condition : Bool;
      sequence_lock : Bool;
   END_VAR
   VAR_TEMP
      cap_detected_tem : Bool;
      sealing_pulse : Bool;
      part_left_sealing : Bool;
   END_VAR
   VAR_TEMP   // added for the SCL form of the ladder/FBD networks
      _w1 : Bool;
      _w2 : Bool;
      _w3 : Bool;
   END_VAR
BEGIN

REGION Network 1: define cretical condition to start the station
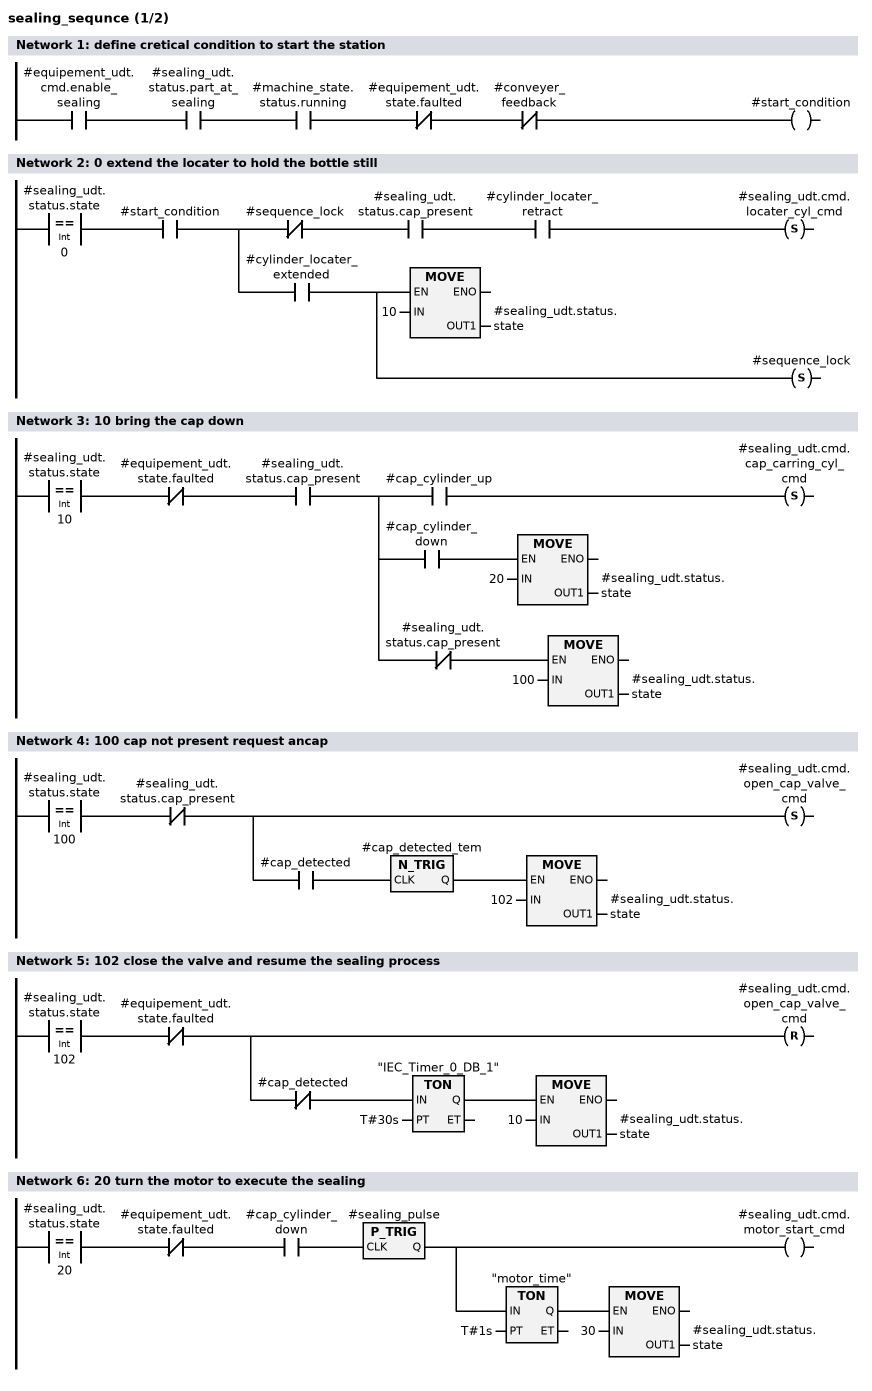
   RUNG wire#powerrail
      Contact( #equipement_udt.cmd.enable_sealing )
      Contact( #sealing_udt.status.part_at_sealing )
      Contact( #machine_state.status.running )
      I_Contact( #equipement_udt.state.faulted )
      I_Contact( #conveyer_feedback )
      Coil( #start_condition )
   END_RUNG
   // the same network as SCL:
   #start_condition := #equipement_udt.cmd.enable_sealing AND #sealing_udt.status.part_at_sealing AND #machine_state.status.running AND NOT #equipement_udt.state.faulted AND NOT #conveyer_feedback;
END_REGION

REGION Network 2: 0 extend the locater to hold the bottle still
   RUNG wire#powerrail
      { S7_Templates := "SrcType := Int" } EQ_Contact(in1 := #sealing_udt.status.state, in2 := 0)
      Contact( #start_condition )
      wire#w1
      I_Contact( #sequence_lock )
      Contact( #sealing_udt.status.cap_present )
      Contact( #cylinder_locater_retract )
      S_Coil( #sealing_udt.cmd.locater_cyl_cmd )
   END_RUNG
   RUNG wire#w1
      Contact( #cylinder_locater_extended )
      wire#w2
      Move(in := 10, out1 => #sealing_udt.status.state)
   END_RUNG
   RUNG wire#w2
      S_Coil( #sequence_lock )
   END_RUNG
   // the same network as SCL:
   #_w1 := (#sealing_udt.status.state = 0) AND #start_condition;
   IF #_w1 AND NOT #sequence_lock AND #sealing_udt.status.cap_present AND #cylinder_locater_retract THEN
       #sealing_udt.cmd.locater_cyl_cmd := TRUE;
   END_IF;
   IF #_w1 AND #cylinder_locater_extended THEN
       #sealing_udt.status.state := 10;
       #sequence_lock := TRUE;
   END_IF;
END_REGION

REGION Network 3: 10 bring the cap down
   RUNG wire#powerrail
      { S7_Templates := "SrcType := Int" } EQ_Contact(in1 := #sealing_udt.status.state, in2 := 10)
      I_Contact( #equipement_udt.state.faulted )
      Contact( #sealing_udt.status.cap_present )
      wire#w1
      Contact( #cap_cylinder_up )
      S_Coil( #sealing_udt.cmd.cap_carring_cyl_cmd )
   END_RUNG
   RUNG wire#w1
      Contact( #cap_cylinder_down )
      Move(in := 20, out1 => #sealing_udt.status.state)
   END_RUNG
   RUNG wire#w1
      I_Contact( #sealing_udt.status.cap_present )
      Move(in := 100, out1 => #sealing_udt.status.state)
   END_RUNG
   // the same network as SCL:
   #_w1 := (#sealing_udt.status.state = 10) AND NOT #equipement_udt.state.faulted AND #sealing_udt.status.cap_present;
   IF #_w1 AND #cap_cylinder_up THEN #sealing_udt.cmd.cap_carring_cyl_cmd := TRUE; END_IF;
   IF #_w1 AND #cap_cylinder_down THEN #sealing_udt.status.state := 20; END_IF;
   IF #_w1 AND NOT #sealing_udt.status.cap_present THEN #sealing_udt.status.state := 100; END_IF;
END_REGION

REGION Network 4: 100 cap not present request ancap
   RUNG wire#powerrail
      { S7_Templates := "SrcType := Int" } EQ_Contact(in1 := #sealing_udt.status.state, in2 := 100)
      I_Contact( #sealing_udt.status.cap_present )
      wire#w1
      S_Coil( #sealing_udt.cmd.open_cap_valve_cmd )
   END_RUNG
   RUNG wire#w1
      Contact( #cap_detected )
      N_Trig( #cap_detected_tem )
      Move(in := 102, out1 => #sealing_udt.status.state)
   END_RUNG
   // the same network as SCL:
   #_w1 := (#sealing_udt.status.state = 100) AND NOT #sealing_udt.status.cap_present;
   IF #_w1 THEN #sealing_udt.cmd.open_cap_valve_cmd := TRUE; END_IF;
   #_w2 := #_w1 AND #cap_detected;
   #_w3 := NOT #_w2 AND #cap_detected_tem;   // falling edge
   #cap_detected_tem := #_w2;
   IF #_w3 THEN #sealing_udt.status.state := 102; END_IF;
END_REGION

REGION Network 5: 102 close the valve and resume the sealing process
   #_w1 := (#sealing_udt.status.state = 102) AND NOT #equipement_udt.state.faulted;
   IF #_w1 THEN #sealing_udt.cmd.open_cap_valve_cmd := FALSE; END_IF;
   "IEC_Timer_0_DB_1".TON(IN := #_w1 AND NOT #cap_detected, PT := T#30s);
   IF "IEC_Timer_0_DB_1".Q THEN #sealing_udt.status.state := 10; END_IF;
END_REGION

REGION Network 6: 20 turn the motor to execute the sealing
   #_w1 := (#sealing_udt.status.state = 20) AND NOT #equipement_udt.state.faulted AND #cap_cylinder_down;
   #_w2 := #_w1 AND NOT #sealing_pulse;   // rising edge
   #sealing_pulse := #_w1;
   #sealing_udt.cmd.motor_start_cmd := #_w2;
   "motor_time".TON(IN := #_w2, PT := T#1s);
   IF "motor_time".Q THEN #sealing_udt.status.state := 30; END_IF;
END_REGION

REGION Network 7: 30 move the cylinder up and locater retracted position
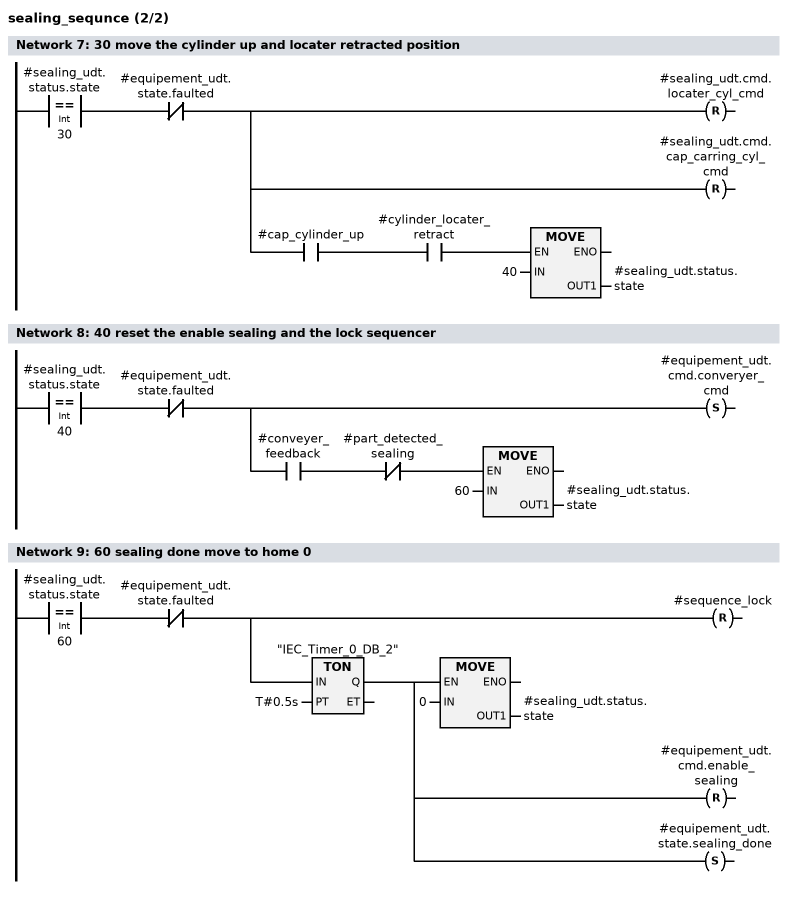
   RUNG wire#powerrail
      { S7_Templates := "SrcType := Int" } EQ_Contact(in1 := #sealing_udt.status.state, in2 := 30)
      I_Contact( #equipement_udt.state.faulted )
      wire#w1
      R_Coil( #sealing_udt.cmd.locater_cyl_cmd )
   END_RUNG
   RUNG wire#w1
      R_Coil( #sealing_udt.cmd.cap_carring_cyl_cmd )
   END_RUNG
   RUNG wire#w1
      Contact( #cap_cylinder_up )
      Contact( #cylinder_locater_retract )
      Move(in := 40, out1 => #sealing_udt.status.state)
   END_RUNG
   // the same network as SCL:
   #_w1 := (#sealing_udt.status.state = 30) AND NOT #equipement_udt.state.faulted;
   IF #_w1 THEN
       #sealing_udt.cmd.locater_cyl_cmd := FALSE;
       #sealing_udt.cmd.cap_carring_cyl_cmd := FALSE;
   END_IF;
   IF #_w1 AND #cap_cylinder_up AND #cylinder_locater_retract THEN #sealing_udt.status.state := 40; END_IF;
END_REGION

REGION Network 8: 40 reset the enable sealing and the lock sequencer
   RUNG wire#powerrail
      { S7_Templates := "SrcType := Int" } EQ_Contact(in1 := #sealing_udt.status.state, in2 := 40)
      I_Contact( #equipement_udt.state.faulted )
      wire#w1
      S_Coil( #equipement_udt.cmd.converyer_cmd )
   END_RUNG
   RUNG wire#w1
      Contact( #conveyer_feedback )
      I_Contact( #part_detected_sealing )
      Move(in := 60, out1 => #sealing_udt.status.state)
   END_RUNG
   // the same network as SCL:
   #_w1 := (#sealing_udt.status.state = 40) AND NOT #equipement_udt.state.faulted;
   IF #_w1 THEN #equipement_udt.cmd.converyer_cmd := TRUE; END_IF;
   IF #_w1 AND #conveyer_feedback AND NOT #part_detected_sealing THEN
       #sealing_udt.status.state := 60;
   END_IF;
END_REGION

REGION Network 9: 60 sealing done move to home 0
   #_w1 := (#sealing_udt.status.state = 60) AND NOT #equipement_udt.state.faulted;
   IF #_w1 THEN #sequence_lock := FALSE; END_IF;
   "IEC_Timer_0_DB_2".TON(IN := #_w1, PT := T#0.5s);
   IF "IEC_Timer_0_DB_2".Q THEN
       #sealing_udt.status.state := 0;
       #equipement_udt.cmd.enable_sealing := FALSE;
       #equipement_udt.state.sealing_done := TRUE;
   END_IF;
END_REGION
END_FUNCTION_BLOCK

FUNCTION "main_capping" : Void   // FC7, LAD
{ S7_Optimized_Access := 'TRUE' }
VERSION : 0.1
BEGIN

REGION Network 1: call generic handler for the capping cylinder locater
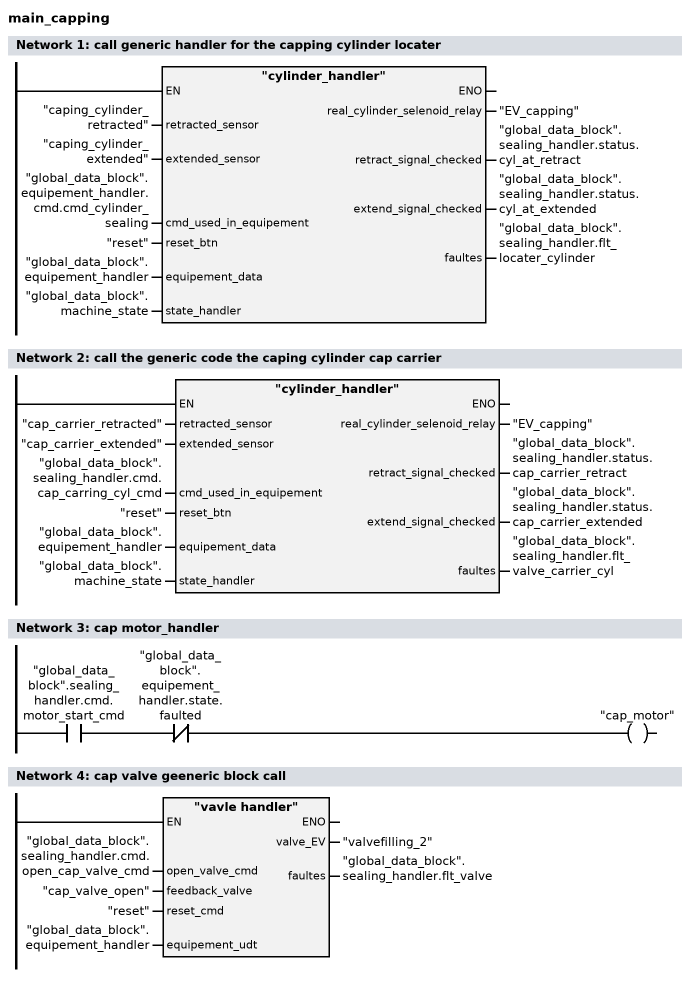
   RUNG wire#powerrail
      "cylinder_handler"(retracted_sensor := "caping_cylinder_retracted", extended_sensor := "caping_cylinder_extended", cmd_used_in_equipement := "global_data_block".equipement_handler.cmd.cmd_cylinder_sealing, reset_btn := "reset", equipement_data := "global_data_block".equipement_handler, state_handler := "global_data_block".machine_state, real_cylinder_selenoid_relay => "EV_capping", retract_signal_checked => "global_data_block".sealing_handler.status.cyl_at_retract, extend_signal_checked => "global_data_block".sealing_handler.status.cyl_at_extended, faultes => "global_data_block".sealing_handler.flt_locater_cylinder)
   END_RUNG
   // the same network as SCL:
   "cylinder_handler"(retracted_sensor := "caping_cylinder_retracted",
                      extended_sensor := "caping_cylinder_extended",
                      cmd_used_in_equipement := "global_data_block".equipement_handler.cmd.cmd_cylinder_sealing,
                      reset_btn := "reset",
                      equipement_data := "global_data_block".equipement_handler,
                      state_handler := "global_data_block".machine_state,
                      real_cylinder_selenoid_relay => "EV_capping",
                      retract_signal_checked => "global_data_block".sealing_handler.status.cyl_at_retract,
                      extend_signal_checked => "global_data_block".sealing_handler.status.cyl_at_extended,
                      faultes => "global_data_block".sealing_handler.flt_locater_cylinder);
END_REGION

REGION Network 2: call the generic code the caping cylinder cap carrier
   RUNG wire#powerrail
      "cylinder_handler"(retracted_sensor := "cap_carrier_retracted", extended_sensor := "cap_carrier_extended", cmd_used_in_equipement := "global_data_block".sealing_handler.cmd.cap_carring_cyl_cmd, reset_btn := "reset", equipement_data := "global_data_block".equipement_handler, state_handler := "global_data_block".machine_state, real_cylinder_selenoid_relay => "EV_capping", retract_signal_checked => "global_data_block".sealing_handler.status.cap_carrier_retract, extend_signal_checked => "global_data_block".sealing_handler.status.cap_carrier_extended, faultes => "global_data_block".sealing_handler.flt_valve_carrier_cyl)
   END_RUNG
   // the same network as SCL:
   "cylinder_handler"(retracted_sensor := "cap_carrier_retracted",
                      extended_sensor := "cap_carrier_extended",
                      cmd_used_in_equipement := "global_data_block".sealing_handler.cmd.cap_carring_cyl_cmd,
                      reset_btn := "reset",
                      equipement_data := "global_data_block".equipement_handler,
                      state_handler := "global_data_block".machine_state,
                      real_cylinder_selenoid_relay => "EV_capping",
                      retract_signal_checked => "global_data_block".sealing_handler.status.cap_carrier_retract,
                      extend_signal_checked => "global_data_block".sealing_handler.status.cap_carrier_extended,
                      faultes => "global_data_block".sealing_handler.flt_valve_carrier_cyl);
END_REGION

REGION Network 3: cap motor_handler
   RUNG wire#powerrail
      Contact( "global_data_block".sealing_handler.cmd.motor_start_cmd )
      I_Contact( "global_data_block".equipement_handler.state.faulted )
      Coil( "cap_motor" )
   END_RUNG
   // the same network as SCL:
   "cap_motor" := "global_data_block".sealing_handler.cmd.motor_start_cmd AND NOT "global_data_block".equipement_handler.state.faulted;
END_REGION

REGION Network 4: cap valve geeneric block call
   RUNG wire#powerrail
      "vavle handler"(open_valve_cmd := "global_data_block".sealing_handler.cmd.open_cap_valve_cmd, feedback_valve := "cap_valve_open", reset_cmd := "reset", equipement_udt := "global_data_block".equipement_handler, valve_EV => "valvefilling_2", faultes => "global_data_block".sealing_handler.flt_valve)
   END_RUNG
   // the same network as SCL:
   "vavle handler"(open_valve_cmd := "global_data_block".sealing_handler.cmd.open_cap_valve_cmd,
                   feedback_valve := "cap_valve_open",
                   reset_cmd := "reset",
                   equipement_udt := "global_data_block".equipement_handler,
                   valve_EV => "valvefilling_2",
                   faultes => "global_data_block".sealing_handler.flt_valve);
END_REGION
END_FUNCTION

// folder: equipement/filling

FUNCTION_BLOCK "filling_sequence"   // FB8, LAD
{ S7_Optimized_Access := 'TRUE' }
VERSION : 0.1
   VAR_INPUT
      conveyer_feedback : Bool;
      part_at_felling : Bool;
      locater_extended : Bool;
      locater_retracted : Bool;
      valve_cylinder_up : Bool;
      valve_cylinder_down : Bool;
   END_VAR
   VAR_IN_OUT
      equipement_data : "udt_equipement";
      state_handler : "udt_state_handler";
      filling_udt : "filling_station_udt";
   END_VAR
   VAR
      sequencer_lock : Bool;
      cycle_condition : Bool;
   END_VAR
   VAR_TEMP
      part_left_filling : Bool;
   END_VAR
   VAR_TEMP   // added for the SCL form of the ladder/FBD networks
      _w1 : Bool;
      _w2 : Bool;
   END_VAR
BEGIN

REGION Network 1: START CONDITION
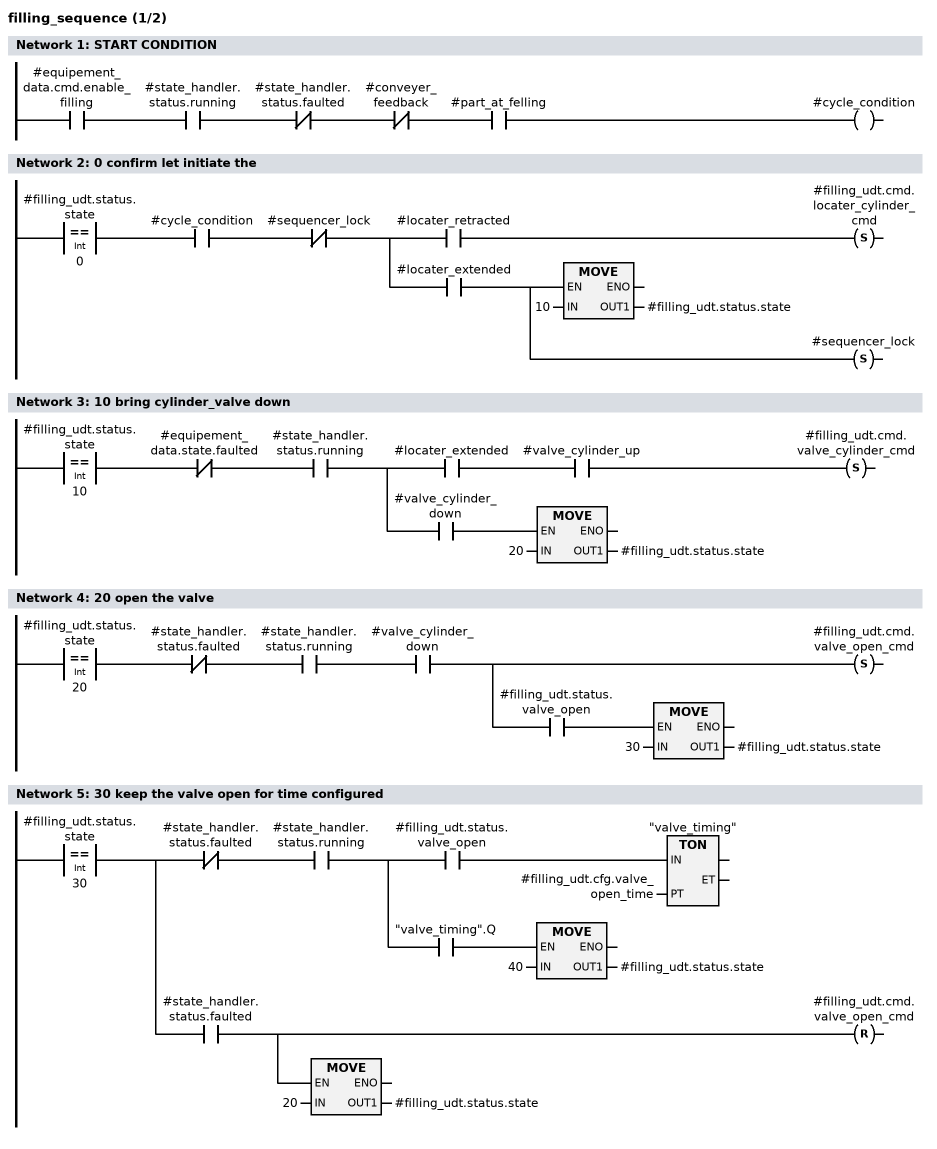
   RUNG wire#powerrail
      Contact( #equipement_data.cmd.enable_filling )
      Contact( #state_handler.status.running )
      I_Contact( #state_handler.status.faulted )
      I_Contact( #conveyer_feedback )
      Contact( #part_at_felling )
      Coil( #cycle_condition )
   END_RUNG
   // the same network as SCL:
   #cycle_condition := #equipement_data.cmd.enable_filling AND #state_handler.status.running AND NOT #state_handler.status.faulted AND NOT #conveyer_feedback AND #part_at_felling;
END_REGION

REGION Network 2: 0 confirm let initiate the
   RUNG wire#powerrail
      { S7_Templates := "SrcType := Int" } EQ_Contact(in1 := #filling_udt.status.state, in2 := 0)
      Contact( #cycle_condition )
      I_Contact( #sequencer_lock )
      wire#w1
      Contact( #locater_retracted )
      S_Coil( #filling_udt.cmd.locater_cylinder_cmd )
   END_RUNG
   RUNG wire#w1
      Contact( #locater_extended )
      wire#w2
      Move(in := 10, out1 => #filling_udt.status.state)
   END_RUNG
   RUNG wire#w2
      S_Coil( #sequencer_lock )
   END_RUNG
   // the same network as SCL:
   #_w1 := (#filling_udt.status.state = 0) AND #cycle_condition AND NOT #sequencer_lock;
   IF #_w1 AND #locater_retracted THEN #filling_udt.cmd.locater_cylinder_cmd := TRUE; END_IF;
   IF #_w1 AND #locater_extended THEN
       #filling_udt.status.state := 10;
       #sequencer_lock := TRUE;
   END_IF;
END_REGION

REGION Network 3: 10 bring cylinder_valve down
   RUNG wire#powerrail
      { S7_Templates := "SrcType := Int" } EQ_Contact(in1 := #filling_udt.status.state, in2 := 10)
      I_Contact( #equipement_data.state.faulted )
      Contact( #state_handler.status.running )
      wire#w1
      Contact( #locater_extended )
      Contact( #valve_cylinder_up )
      S_Coil( #filling_udt.cmd.valve_cylinder_cmd )
   END_RUNG
   RUNG wire#w1
      Contact( #valve_cylinder_down )
      Move(in := 20, out1 => #filling_udt.status.state)
   END_RUNG
   // the same network as SCL:
   #_w1 := (#filling_udt.status.state = 10) AND NOT #equipement_data.state.faulted AND #state_handler.status.running;
   IF #_w1 AND #locater_extended AND #valve_cylinder_up THEN
       #filling_udt.cmd.valve_cylinder_cmd := TRUE;
   END_IF;
   IF #_w1 AND #valve_cylinder_down THEN #filling_udt.status.state := 20; END_IF;
END_REGION

REGION Network 4: 20 open the valve
   RUNG wire#powerrail
      { S7_Templates := "SrcType := Int" } EQ_Contact(in1 := #filling_udt.status.state, in2 := 20)
      I_Contact( #state_handler.status.faulted )
      Contact( #state_handler.status.running )
      Contact( #valve_cylinder_down )
      wire#w1
      S_Coil( #filling_udt.cmd.valve_open_cmd )
   END_RUNG
   RUNG wire#w1
      Contact( #filling_udt.status.valve_open )
      Move(in := 30, out1 => #filling_udt.status.state)
   END_RUNG
   // the same network as SCL:
   #_w1 := (#filling_udt.status.state = 20) AND NOT #state_handler.status.faulted AND #state_handler.status.running AND #valve_cylinder_down;
   IF #_w1 THEN #filling_udt.cmd.valve_open_cmd := TRUE; END_IF;
   IF #_w1 AND #filling_udt.status.valve_open THEN #filling_udt.status.state := 30; END_IF;
END_REGION

REGION Network 5: 30 keep the valve open for time configured
   #_w1 := #filling_udt.status.state = 30;
   #_w2 := #_w1 AND NOT #state_handler.status.faulted AND #state_handler.status.running;
   "valve_timing".TON(IN := #_w2 AND #filling_udt.status.valve_open, PT := #filling_udt.cfg.valve_open_time);
   IF #_w2 AND "valve_timing".Q THEN #filling_udt.status.state := 40; END_IF;
   IF #_w1 AND #state_handler.status.faulted THEN
       #filling_udt.cmd.valve_open_cmd := FALSE;
       #filling_udt.status.state := 20;
   END_IF;
END_REGION

REGION Network 6: 40 retract the locater
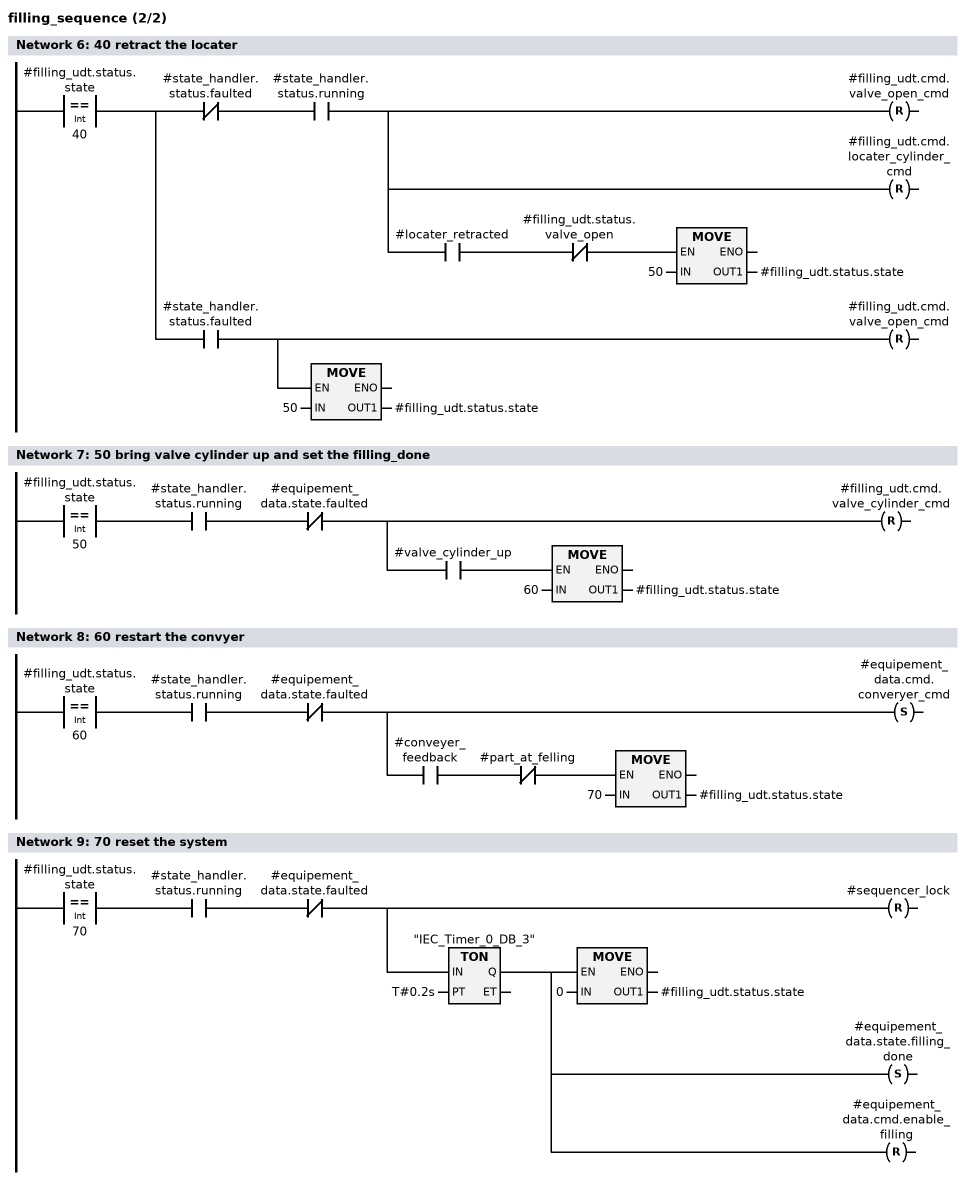
   RUNG wire#powerrail
      { S7_Templates := "SrcType := Int" } EQ_Contact(in1 := #filling_udt.status.state, in2 := 40)
      wire#w1
      I_Contact( #state_handler.status.faulted )
      Contact( #state_handler.status.running )
      wire#w2
      R_Coil( #filling_udt.cmd.valve_open_cmd )
   END_RUNG
   RUNG wire#w2
      R_Coil( #filling_udt.cmd.locater_cylinder_cmd )
   END_RUNG
   RUNG wire#w2
      Contact( #locater_retracted )
      I_Contact( #filling_udt.status.valve_open )
      Move(in := 50, out1 => #filling_udt.status.state)
   END_RUNG
   RUNG wire#w1
      Contact( #state_handler.status.faulted )
      wire#w3
      R_Coil( #filling_udt.cmd.valve_open_cmd )
   END_RUNG
   RUNG wire#w3
      Move(in := 50, out1 => #filling_udt.status.state)
   END_RUNG
   // the same network as SCL:
   #_w1 := #filling_udt.status.state = 40;
   #_w2 := #_w1 AND NOT #state_handler.status.faulted AND #state_handler.status.running;
   IF #_w2 THEN
       #filling_udt.cmd.valve_open_cmd := FALSE;
       #filling_udt.cmd.locater_cylinder_cmd := FALSE;
   END_IF;
   IF #_w2 AND #locater_retracted AND NOT #filling_udt.status.valve_open THEN
       #filling_udt.status.state := 50;
   END_IF;
   IF #_w1 AND #state_handler.status.faulted THEN
       #filling_udt.cmd.valve_open_cmd := FALSE;
       #filling_udt.status.state := 50;
   END_IF;
END_REGION

REGION Network 7: 50 bring valve cylinder up and set the filling_done
   RUNG wire#powerrail
      { S7_Templates := "SrcType := Int" } EQ_Contact(in1 := #filling_udt.status.state, in2 := 50)
      Contact( #state_handler.status.running )
      I_Contact( #equipement_data.state.faulted )
      wire#w1
      R_Coil( #filling_udt.cmd.valve_cylinder_cmd )
   END_RUNG
   RUNG wire#w1
      Contact( #valve_cylinder_up )
      Move(in := 60, out1 => #filling_udt.status.state)
   END_RUNG
   // the same network as SCL:
   #_w1 := (#filling_udt.status.state = 50) AND #state_handler.status.running AND NOT #equipement_data.state.faulted;
   IF #_w1 THEN #filling_udt.cmd.valve_cylinder_cmd := FALSE; END_IF;
   IF #_w1 AND #valve_cylinder_up THEN #filling_udt.status.state := 60; END_IF;
END_REGION

REGION Network 8: 60 restart the convyer
   RUNG wire#powerrail
      { S7_Templates := "SrcType := Int" } EQ_Contact(in1 := #filling_udt.status.state, in2 := 60)
      Contact( #state_handler.status.running )
      I_Contact( #equipement_data.state.faulted )
      wire#w1
      S_Coil( #equipement_data.cmd.converyer_cmd )
   END_RUNG
   RUNG wire#w1
      Contact( #conveyer_feedback )
      I_Contact( #part_at_felling )
      Move(in := 70, out1 => #filling_udt.status.state)
   END_RUNG
   // the same network as SCL:
   #_w1 := (#filling_udt.status.state = 60) AND #state_handler.status.running AND NOT #equipement_data.state.faulted;
   IF #_w1 THEN #equipement_data.cmd.converyer_cmd := TRUE; END_IF;
   IF #_w1 AND #conveyer_feedback AND NOT #part_at_felling THEN #filling_udt.status.state := 70; END_IF;
END_REGION

REGION Network 9: 70 reset the system
   #_w1 := (#filling_udt.status.state = 70) AND #state_handler.status.running AND NOT #equipement_data.state.faulted;
   IF #_w1 THEN #sequencer_lock := FALSE; END_IF;
   "IEC_Timer_0_DB_3".TON(IN := #_w1, PT := T#0.2s);
   IF "IEC_Timer_0_DB_3".Q THEN
       #filling_udt.status.state := 0;
       #equipement_data.state.filling_done := TRUE;
       #equipement_data.cmd.enable_filling := FALSE;
   END_IF;
END_REGION
END_FUNCTION_BLOCK

FUNCTION "main_filling" : Void   // FC6, LAD
{ S7_Optimized_Access := 'TRUE' }
VERSION : 0.1
BEGIN

REGION Network 1: call generic code to handle locater cylinder befaviours
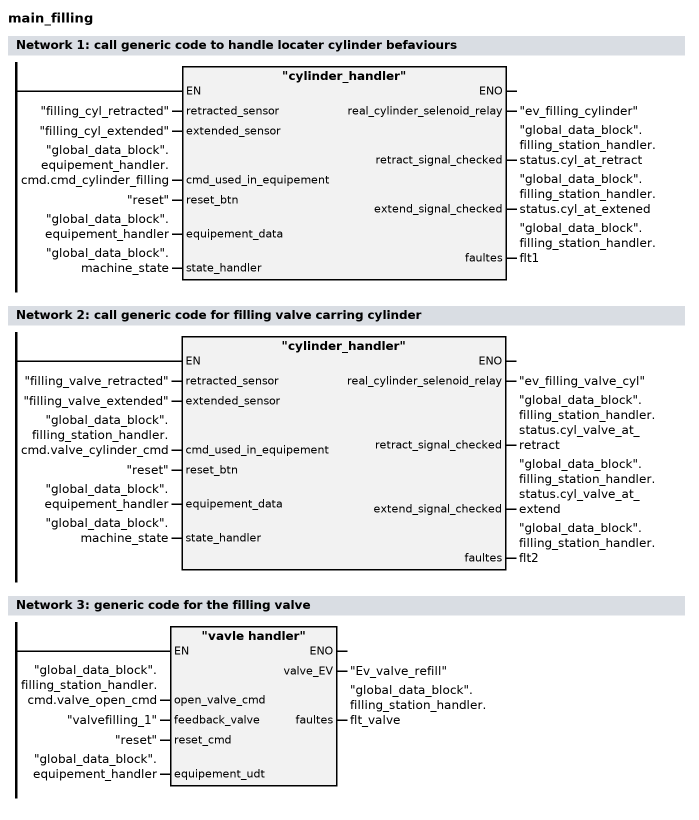
   RUNG wire#powerrail
      "cylinder_handler"(retracted_sensor := "filling_cyl_retracted", extended_sensor := "filling_cyl_extended", cmd_used_in_equipement := "global_data_block".equipement_handler.cmd.cmd_cylinder_filling, reset_btn := "reset", equipement_data := "global_data_block".equipement_handler, state_handler := "global_data_block".machine_state, real_cylinder_selenoid_relay => "ev_filling_cylinder", retract_signal_checked => "global_data_block".filling_station_handler.status.cyl_at_retract, extend_signal_checked => "global_data_block".filling_station_handler.status.cyl_at_extened, faultes => "global_data_block".filling_station_handler.flt1)
   END_RUNG
   // the same network as SCL:
   "cylinder_handler"(retracted_sensor := "filling_cyl_retracted",
                      extended_sensor := "filling_cyl_extended",
                      cmd_used_in_equipement := "global_data_block".equipement_handler.cmd.cmd_cylinder_filling,
                      reset_btn := "reset",
                      equipement_data := "global_data_block".equipement_handler,
                      state_handler := "global_data_block".machine_state,
                      real_cylinder_selenoid_relay => "ev_filling_cylinder",
                      retract_signal_checked => "global_data_block".filling_station_handler.status.cyl_at_retract,
                      extend_signal_checked => "global_data_block".filling_station_handler.status.cyl_at_extened,
                      faultes => "global_data_block".filling_station_handler.flt1);
END_REGION

REGION Network 2: call generic code for filling valve carring cylinder
   RUNG wire#powerrail
      "cylinder_handler"(retracted_sensor := "filling_valve_retracted", extended_sensor := "filling_valve_extended", cmd_used_in_equipement := "global_data_block".filling_station_handler.cmd.valve_cylinder_cmd, reset_btn := "reset", equipement_data := "global_data_block".equipement_handler, state_handler := "global_data_block".machine_state, real_cylinder_selenoid_relay => "ev_filling_valve_cyl", retract_signal_checked => "global_data_block".filling_station_handler.status.cyl_valve_at_retract, extend_signal_checked => "global_data_block".filling_station_handler.status.cyl_valve_at_extend, faultes => "global_data_block".filling_station_handler.flt2)
   END_RUNG
   // the same network as SCL:
   "cylinder_handler"(retracted_sensor := "filling_valve_retracted",
                      extended_sensor := "filling_valve_extended",
                      cmd_used_in_equipement := "global_data_block".filling_station_handler.cmd.valve_cylinder_cmd,
                      reset_btn := "reset",
                      equipement_data := "global_data_block".equipement_handler,
                      state_handler := "global_data_block".machine_state,
                      real_cylinder_selenoid_relay => "ev_filling_valve_cyl",
                      retract_signal_checked => "global_data_block".filling_station_handler.status.cyl_valve_at_retract,
                      extend_signal_checked => "global_data_block".filling_station_handler.status.cyl_valve_at_extend,
                      faultes => "global_data_block".filling_station_handler.flt2);
END_REGION

REGION Network 3: generic code for the filling valve
   RUNG wire#powerrail
      "vavle handler"(open_valve_cmd := "global_data_block".filling_station_handler.cmd.valve_open_cmd, feedback_valve := "valvefilling_1", reset_cmd := "reset", equipement_udt := "global_data_block".equipement_handler, valve_EV => "Ev_valve_refill", faultes => "global_data_block".filling_station_handler.flt_valve)
   END_RUNG
   // the same network as SCL:
   "vavle handler"(open_valve_cmd := "global_data_block".filling_station_handler.cmd.valve_open_cmd,
                   feedback_valve := "valvefilling_1",
                   reset_cmd := "reset",
                   equipement_udt := "global_data_block".equipement_handler,
                   valve_EV => "Ev_valve_refill",
                   faultes => "global_data_block".filling_station_handler.flt_valve);
END_REGION
END_FUNCTION

// folder: equipement/functions

FUNCTION "scale_function" : Void   // FC3, LAD
{ S7_Optimized_Access := 'TRUE' }
VERSION : 0.1
   VAR_INPUT
      actual_weight_card : Int;
   END_VAR
   VAR_IN_OUT
      scaling_handler : "scaling_udt";
   END_VAR
   VAR_TEMP
      normalised_value : Real;
   END_VAR
BEGIN

REGION Network 1: normalize the hardward readings
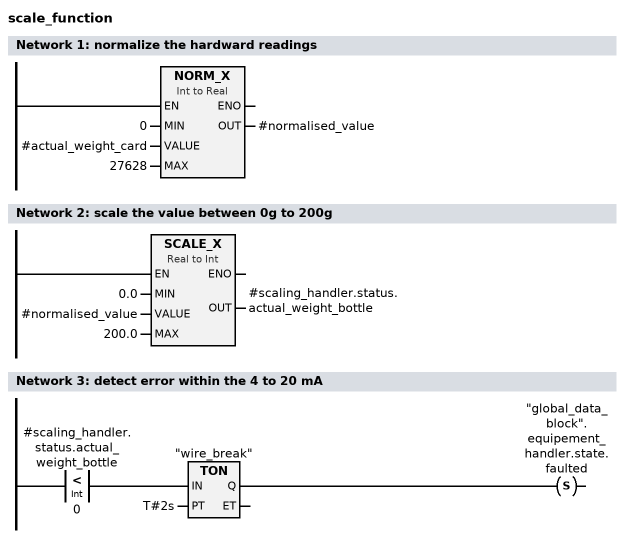
   RUNG wire#powerrail
      { S7_Templates := "[SrcType := Int, DestType := Real]" } Normalize(min := 0, value := #actual_weight_card, max := 27628, out => #normalised_value)
   END_RUNG
   // the same network as SCL:
   #normalised_value := NORM_X(MIN := 0, VALUE := #actual_weight_card, MAX := 27628);
END_REGION

REGION Network 2: scale the value between 0g to 200g
   RUNG wire#powerrail
      { S7_Templates := "[SrcType := Real, DestType := Int]" } Scale(min := 0.0, value := #normalised_value, max := 200.0, out => #scaling_handler.status.actual_weight_bottle)
   END_RUNG
   // the same network as SCL:
   #scaling_handler.status.actual_weight_bottle := SCALE_X(MIN := 0.0, VALUE := #normalised_value, MAX := 200.0);
END_REGION

REGION Network 3: detect error within the 4 to 20 mA
   "wire_break".TON(IN := #scaling_handler.status.actual_weight_bottle < 0, PT := T#2s);
   IF "wire_break".Q THEN "global_data_block".equipement_handler.state.faulted := TRUE; END_IF;
END_REGION
END_FUNCTION

FUNCTION "cylinder_handler" : Void   // FC4, LAD
{ S7_Optimized_Access := 'TRUE' }
VERSION : 0.1
   VAR_INPUT
      retracted_sensor : Bool;
      extended_sensor : Bool;
      cmd_used_in_equipement : Bool;
      reset_btn : Bool;
   END_VAR
   VAR_OUTPUT
      real_cylinder_selenoid_relay : Bool;
      retract_signal_checked : Bool;
      extend_signal_checked : Bool;
      faultes : Word;
   END_VAR
   VAR_IN_OUT
      equipement_data : "udt_equipement";
      state_handler : "udt_state_handler";
   END_VAR
   VAR_TEMP
      reset_pulse : Bool;
   END_VAR
   VAR_TEMP   // added for the SCL form of the ladder/FBD networks
      _w1 : Bool;
      _w2 : Bool;
   END_VAR
BEGIN

REGION Network 1: confirm signal from sensors
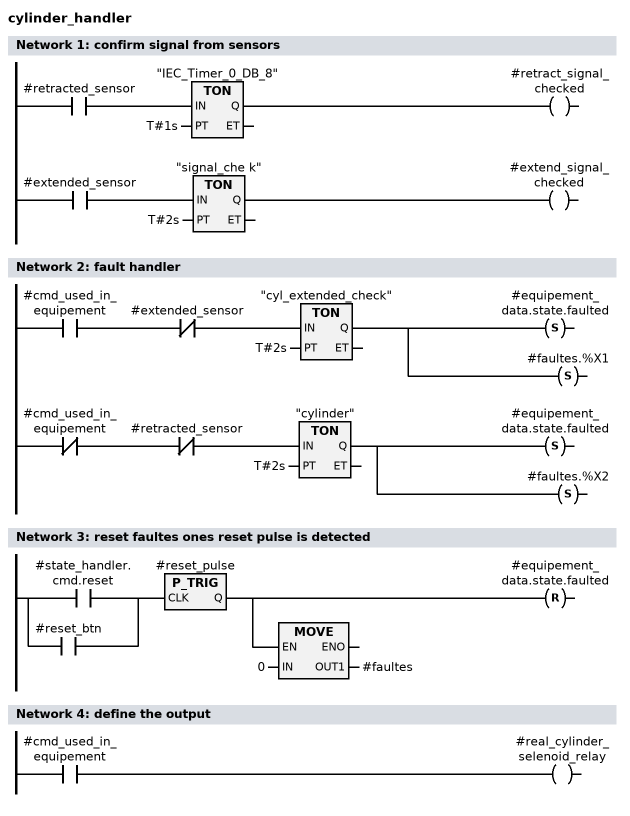
   "IEC_Timer_0_DB_8".TON(IN := #retracted_sensor, PT := T#1s);
   #retract_signal_checked := "IEC_Timer_0_DB_8".Q;
   "signal_che k".TON(IN := #extended_sensor, PT := T#2s);
   #extend_signal_checked := "signal_che k".Q;
END_REGION

REGION Network 2: fault handler
   "cyl_extended_check".TON(IN := #cmd_used_in_equipement AND NOT #extended_sensor, PT := T#2s);
   IF "cyl_extended_check".Q THEN
       #equipement_data.state.faulted := TRUE;
       #faultes.%X1 := TRUE;
   END_IF;
   "cylinder".TON(IN := NOT #cmd_used_in_equipement AND NOT #retracted_sensor, PT := T#2s);
   IF "cylinder".Q THEN
       #equipement_data.state.faulted := TRUE;
       #faultes.%X2 := TRUE;
   END_IF;
END_REGION

REGION Network 3: reset faultes ones reset pulse is detected
   RUNG wire#powerrail
      Contact( #state_handler.cmd.reset )
      wire#w1
      P_Trig( #reset_pulse )
      wire#w2
      R_Coil( #equipement_data.state.faulted )
   END_RUNG
   RUNG wire#powerrail
      Contact( #reset_btn )
   END_RUNG wire#w1
   RUNG wire#w2
      Move(in := 0, out1 => #faultes)
   END_RUNG
   // the same network as SCL:
   #_w1 := #state_handler.cmd.reset OR #reset_btn;
   #_w2 := #_w1 AND NOT #reset_pulse;   // rising edge
   #reset_pulse := #_w1;
   IF #_w2 THEN
       #equipement_data.state.faulted := FALSE;
       #faultes := 0;
   END_IF;
END_REGION

REGION Network 4: define the output
   RUNG wire#powerrail
      Contact( #cmd_used_in_equipement )
      Coil( #real_cylinder_selenoid_relay )
   END_RUNG
   // the same network as SCL:
   #real_cylinder_selenoid_relay := #cmd_used_in_equipement;
END_REGION
END_FUNCTION

FUNCTION "motor_vfd" : Void   // FC5, LAD
{ S7_Optimized_Access := 'TRUE' }
VERSION : 0.1
   VAR_INPUT
      vfd_current_speed : Word;
      "op_set_giving_point(%)" : Int;
      feedback_running : Bool;
      reset : Bool;
      motor_cmd_turn_on : Bool;
   END_VAR
   VAR_OUTPUT
      running : Bool;
      vfd_setpoint : Int;
      faulted : Bool;
      set_point_valid : Bool;
   END_VAR
   VAR_IN_OUT
      equipement_udt : "udt_equipement";
      state_handler : "udt_state_handler";
      vfd_cmd : "vfd_cmd";
      vfd_udt_status : "udt_vfd_status";
   END_VAR
   VAR_TEMP
      reset_pulse : Bool;
   END_VAR
   VAR_TEMP   // added for the SCL form of the ladder/FBD networks
      _w1 : Bool;
      _w2 : Bool;
   END_VAR
BEGIN

REGION Network 1: 1: check setpoint for coherence and consistency
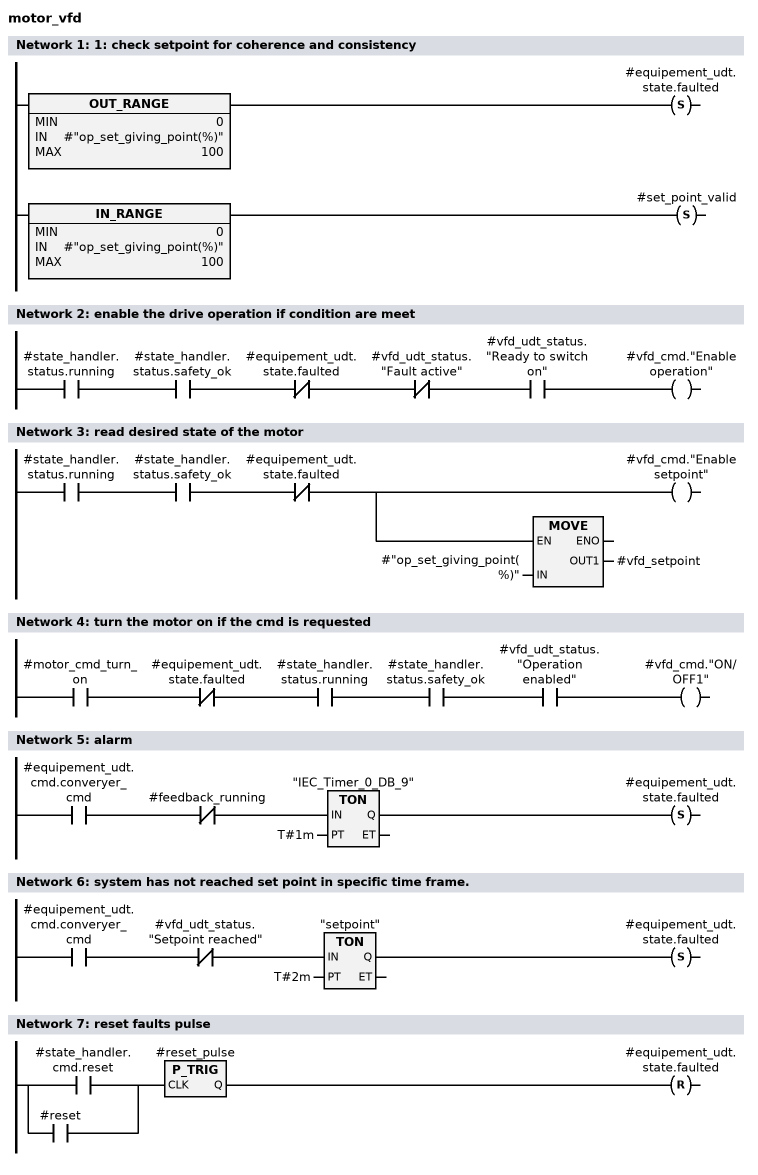
   IF (#"op_set_giving_point(%)" < 0) OR (#"op_set_giving_point(%)" > 100) THEN
       #equipement_udt.state.faulted := TRUE;
   END_IF;
   IF (0 <= #"op_set_giving_point(%)") AND (#"op_set_giving_point(%)" <= 100) THEN
       #set_point_valid := TRUE;
   END_IF;
END_REGION

REGION Network 2: enable the drive operation if condition are meet
   RUNG wire#powerrail
      Contact( #state_handler.status.running )
      Contact( #state_handler.status.safety_ok )
      I_Contact( #equipement_udt.state.faulted )
      I_Contact( #vfd_udt_status."Fault active" )
      Contact( #vfd_udt_status."Ready to switch on" )
      Coil( #vfd_cmd."Enable operation" )
   END_RUNG
   // the same network as SCL:
   #vfd_cmd."Enable operation" := #state_handler.status.running AND #state_handler.status.safety_ok AND NOT #equipement_udt.state.faulted AND NOT #vfd_udt_status."Fault active" AND #vfd_udt_status."Ready to switch on";
END_REGION

REGION Network 3: read desired state of the motor
   RUNG wire#powerrail
      Contact( #state_handler.status.running )
      Contact( #state_handler.status.safety_ok )
      I_Contact( #equipement_udt.state.faulted )
      wire#w1
      Coil( #vfd_cmd."Enable setpoint" )
   END_RUNG
   RUNG wire#w1
      Move(in := #"op_set_giving_point(%)", out1 => #vfd_setpoint)
   END_RUNG
   // the same network as SCL:
   #vfd_cmd."Enable setpoint" := #state_handler.status.running AND #state_handler.status.safety_ok AND NOT #equipement_udt.state.faulted;
   IF #vfd_cmd."Enable setpoint" THEN #vfd_setpoint := #"op_set_giving_point(%)"; END_IF;
END_REGION

REGION Network 4: turn the motor on if the cmd is requested
   RUNG wire#powerrail
      Contact( #motor_cmd_turn_on )
      I_Contact( #equipement_udt.state.faulted )
      Contact( #state_handler.status.running )
      Contact( #state_handler.status.safety_ok )
      Contact( #vfd_udt_status."Operation enabled" )
      Coil( #vfd_cmd."ON/OFF1" )
   END_RUNG
   // the same network as SCL:
   #vfd_cmd."ON/OFF1" := #motor_cmd_turn_on AND NOT #equipement_udt.state.faulted AND #state_handler.status.running AND #state_handler.status.safety_ok AND #vfd_udt_status."Operation enabled";
END_REGION

REGION Network 5: alarm
   "IEC_Timer_0_DB_9".TON(IN := #equipement_udt.cmd.converyer_cmd AND NOT #feedback_running, PT := T#1m);
   IF "IEC_Timer_0_DB_9".Q THEN #equipement_udt.state.faulted := TRUE; END_IF;
END_REGION

REGION Network 6: system has not reached set point in specific time frame.
   "setpoint".TON(IN := #equipement_udt.cmd.converyer_cmd AND NOT #vfd_udt_status."Setpoint reached",
                  PT := T#2m);
   IF "setpoint".Q THEN #equipement_udt.state.faulted := TRUE; END_IF;
END_REGION

REGION Network 7: reset faults pulse
   RUNG wire#powerrail
      Contact( #state_handler.cmd.reset )
      wire#w1
      P_Trig( #reset_pulse )
      R_Coil( #equipement_udt.state.faulted )
   END_RUNG
   RUNG wire#powerrail
      Contact( #reset )
   END_RUNG wire#w1
   // the same network as SCL:
   #_w1 := #state_handler.cmd.reset OR #reset;
   #_w2 := #_w1 AND NOT #reset_pulse;   // rising edge
   #reset_pulse := #_w1;
   IF #_w2 THEN #equipement_udt.state.faulted := FALSE; END_IF;
END_REGION
END_FUNCTION

FUNCTION "vavle handler" : Void   // FC9, LAD
{ S7_Optimized_Access := 'TRUE' }
VERSION : 0.1
   VAR_INPUT
      open_valve_cmd : Bool;
      feedback_valve : Bool;
      reset_cmd : Bool;
   END_VAR
   VAR_OUTPUT
      valve_EV : Bool;
      faultes : Word;
   END_VAR
   VAR_IN_OUT
      equipement_udt : "udt_equipement";
   END_VAR
   VAR_TEMP
      reset_pulse : Bool;
   END_VAR
   VAR_TEMP   // added for the SCL form of the ladder/FBD networks
      _w1 : Bool;
   END_VAR
BEGIN

REGION Network 1: cmd signal check
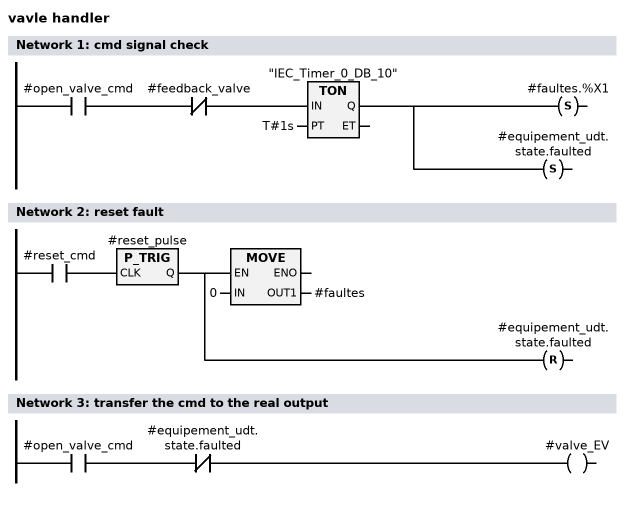
   "IEC_Timer_0_DB_10".TON(IN := #open_valve_cmd AND NOT #feedback_valve, PT := T#1s);
   IF "IEC_Timer_0_DB_10".Q THEN
       #faultes.%X1 := TRUE;
       #equipement_udt.state.faulted := TRUE;
   END_IF;
END_REGION

REGION Network 2: reset fault
   RUNG wire#powerrail
      Contact( #reset_cmd )
      P_Trig( #reset_pulse )
      wire#w1
      Move(in := 0, out1 => #faultes)
   END_RUNG
   RUNG wire#w1
      R_Coil( #equipement_udt.state.faulted )
   END_RUNG
   // the same network as SCL:
   #_w1 := #reset_cmd AND NOT #reset_pulse;   // rising edge
   #reset_pulse := #reset_cmd;
   IF #_w1 THEN
       #faultes := 0;
       #equipement_udt.state.faulted := FALSE;
   END_IF;
END_REGION

REGION Network 3: transfer the cmd to the real output
   RUNG wire#powerrail
      Contact( #open_valve_cmd )
      I_Contact( #equipement_udt.state.faulted )
      Coil( #valve_EV )
   END_RUNG
   // the same network as SCL:
   #valve_EV := #open_valve_cmd AND NOT #equipement_udt.state.faulted;
END_REGION
END_FUNCTION

// folder: equipement/reject

FUNCTION_BLOCK "reject_main"   // FB12, LAD
{ S7_Optimized_Access := 'TRUE' }
VERSION : 0.1
   VAR_INPUT
      part_has_been_rejected : Bool;
      cyl_retracted : Bool;
      part_at_reject : Bool;
      conveyer_feedback : Bool;
      cyl_extended : Bool;
   END_VAR
   VAR_IN_OUT
      state_handler : "udt_state_handler";
      equipement_management : "udt_equipement";
      verification_feedback : "scaling_udt";
      reject_udt : "reject_udt";
   END_VAR
   VAR
      start_condition_1 : Bool;
      repetition_count : Int;
      ton_repetition : TON_TIME;
      increment : Bool;
      reption_enable : Bool;
   END_VAR
   VAR_TEMP
      lock_sequencer : Bool;
      leaving : Bool;
   END_VAR
   VAR_TEMP   // added for the SCL form of the ladder/FBD networks
      _w1 : Bool;
      _w2 : Bool;
      _w3 : Bool;
   END_VAR
BEGIN

REGION Network 1: define the start condition
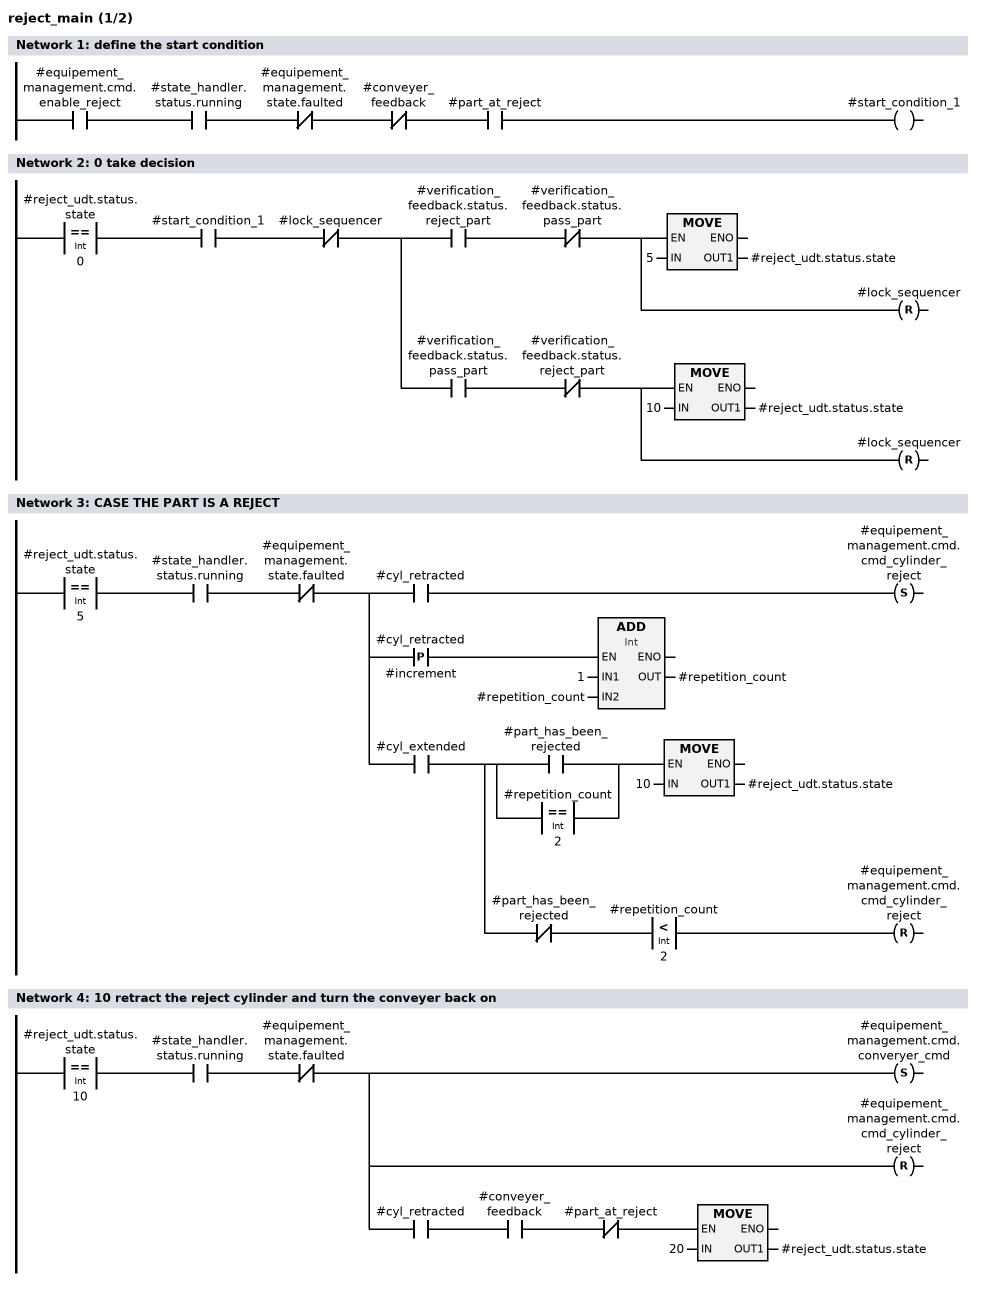
   RUNG wire#powerrail
      Contact( #equipement_management.cmd.enable_reject )
      Contact( #state_handler.status.running )
      I_Contact( #equipement_management.state.faulted )
      I_Contact( #conveyer_feedback )
      Contact( #part_at_reject )
      Coil( #start_condition_1 )
   END_RUNG
   // the same network as SCL:
   #start_condition_1 := #equipement_management.cmd.enable_reject AND #state_handler.status.running AND NOT #equipement_management.state.faulted AND NOT #conveyer_feedback AND #part_at_reject;
END_REGION

REGION Network 2: 0 take decision
   RUNG wire#powerrail
      { S7_Templates := "SrcType := Int" } EQ_Contact(in1 := #reject_udt.status.state, in2 := 0)
      Contact( #start_condition_1 )
      I_Contact( #lock_sequencer )
      wire#w1
      Contact( #verification_feedback.status.reject_part )
      I_Contact( #verification_feedback.status.pass_part )
      wire#w2
      Move(in := 5, out1 => #reject_udt.status.state)
   END_RUNG
   RUNG wire#w2
      R_Coil( #lock_sequencer )
   END_RUNG
   RUNG wire#w1
      Contact( #verification_feedback.status.pass_part )
      I_Contact( #verification_feedback.status.reject_part )
      wire#w3
      Move(in := 10, out1 => #reject_udt.status.state)
   END_RUNG
   RUNG wire#w3
      R_Coil( #lock_sequencer )
   END_RUNG
   // the same network as SCL:
   #_w1 := (#reject_udt.status.state = 0) AND #start_condition_1 AND NOT #lock_sequencer;
   IF #_w1 AND #verification_feedback.status.reject_part AND NOT #verification_feedback.status.pass_part THEN
       #reject_udt.status.state := 5;
       #lock_sequencer := FALSE;
   END_IF;
   IF #_w1 AND #verification_feedback.status.pass_part AND NOT #verification_feedback.status.reject_part THEN
       #reject_udt.status.state := 10;
       #lock_sequencer := FALSE;
   END_IF;
END_REGION

REGION Network 3: CASE THE PART IS A REJECT
   RUNG wire#powerrail
      { S7_Templates := "SrcType := Int" } EQ_Contact(in1 := #reject_udt.status.state, in2 := 5)
      Contact( #state_handler.status.running )
      I_Contact( #equipement_management.state.faulted )
      wire#w1
      Contact( #cyl_retracted )
      S_Coil( #equipement_management.cmd.cmd_cylinder_reject )
   END_RUNG
   RUNG wire#w1
      P_Contact(operand := #cyl_retracted, bit := #increment)
      { S7_Templates := "SrcType := Int" } Add(in1 := 1, in2 := #repetition_count, out => #repetition_count)
   END_RUNG
   RUNG wire#w1
      Contact( #cyl_extended )
      wire#w2
      Contact( #part_has_been_rejected )
      wire#w3
      Move(in := 10, out1 => #reject_udt.status.state)
   END_RUNG
   RUNG wire#w2
      { S7_Templates := "SrcType := Int" } EQ_Contact(in1 := #repetition_count, in2 := 2)
   END_RUNG wire#w3
   RUNG wire#w2
      I_Contact( #part_has_been_rejected )
      { S7_Templates := "SrcType := Int" } LT_Contact(in1 := #repetition_count, in2 := 2)
      R_Coil( #equipement_management.cmd.cmd_cylinder_reject )
   END_RUNG
   // the same network as SCL:
   #_w1 := (#reject_udt.status.state = 5) AND #state_handler.status.running AND NOT #equipement_management.state.faulted;
   IF #_w1 AND #cyl_retracted THEN #equipement_management.cmd.cmd_cylinder_reject := TRUE; END_IF;
   #_w2 := #_w1 AND #cyl_retracted AND NOT #increment;   // rising edge of #cyl_retracted
   #increment := #cyl_retracted;
   IF #_w2 THEN #repetition_count := 1 + #repetition_count; END_IF;
   #_w3 := #_w1 AND #cyl_extended;
   IF #_w3 AND (#part_has_been_rejected OR (#repetition_count = 2)) THEN
       #reject_udt.status.state := 10;
   END_IF;
   IF #_w3 AND NOT #part_has_been_rejected AND (#repetition_count < 2) THEN
       #equipement_management.cmd.cmd_cylinder_reject := FALSE;
   END_IF;
END_REGION

REGION Network 4: 10 retract the reject cylinder and turn the conveyer back on
   RUNG wire#powerrail
      { S7_Templates := "SrcType := Int" } EQ_Contact(in1 := #reject_udt.status.state, in2 := 10)
      Contact( #state_handler.status.running )
      I_Contact( #equipement_management.state.faulted )
      wire#w1
      S_Coil( #equipement_management.cmd.converyer_cmd )
   END_RUNG
   RUNG wire#w1
      R_Coil( #equipement_management.cmd.cmd_cylinder_reject )
   END_RUNG
   RUNG wire#w1
      Contact( #cyl_retracted )
      Contact( #conveyer_feedback )
      I_Contact( #part_at_reject )
      Move(in := 20, out1 => #reject_udt.status.state)
   END_RUNG
   // the same network as SCL:
   #_w1 := (#reject_udt.status.state = 10) AND #state_handler.status.running AND NOT #equipement_management.state.faulted;
   IF #_w1 THEN
       #equipement_management.cmd.converyer_cmd := TRUE;
       #equipement_management.cmd.cmd_cylinder_reject := FALSE;
   END_IF;
   IF #_w1 AND #cyl_retracted AND #conveyer_feedback AND NOT #part_at_reject THEN
       #reject_udt.status.state := 20;
   END_IF;
END_REGION

REGION Network 5: 20 disable the reject enable and allow for more part
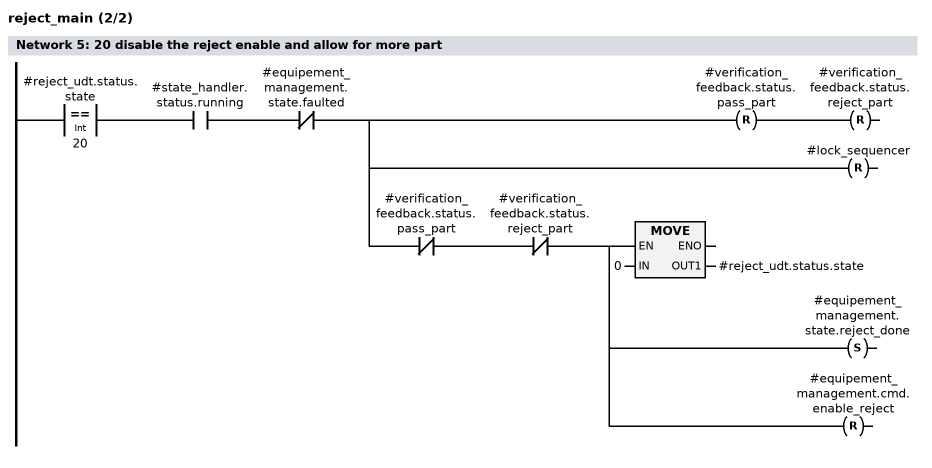
   RUNG wire#powerrail
      { S7_Templates := "SrcType := Int" } EQ_Contact(in1 := #reject_udt.status.state, in2 := 20)
      Contact( #state_handler.status.running )
      I_Contact( #equipement_management.state.faulted )
      wire#w1
      R_Coil( #verification_feedback.status.pass_part )
      R_Coil( #verification_feedback.status.reject_part )
   END_RUNG
   RUNG wire#w1
      R_Coil( #lock_sequencer )
   END_RUNG
   RUNG wire#w1
      I_Contact( #verification_feedback.status.pass_part )
      I_Contact( #verification_feedback.status.reject_part )
      wire#w2
      Move(in := 0, out1 => #reject_udt.status.state)
   END_RUNG
   RUNG wire#w2
      S_Coil( #equipement_management.state.reject_done )
   END_RUNG
   RUNG wire#w2
      R_Coil( #equipement_management.cmd.enable_reject )
   END_RUNG
   // the same network as SCL:
   #_w1 := (#reject_udt.status.state = 20) AND #state_handler.status.running AND NOT #equipement_management.state.faulted;
   IF #_w1 THEN
       #verification_feedback.status.pass_part := FALSE;
       #verification_feedback.status.reject_part := FALSE;
       #lock_sequencer := FALSE;
   END_IF;
   IF #_w1 AND NOT #verification_feedback.status.pass_part AND NOT #verification_feedback.status.reject_part THEN
       #reject_udt.status.state := 0;
       #equipement_management.state.reject_done := TRUE;
       #equipement_management.cmd.enable_reject := FALSE;
   END_IF;
END_REGION
END_FUNCTION_BLOCK

FUNCTION "main_reject" : Void   // FC8, LAD
{ S7_Optimized_Access := 'TRUE' }
VERSION : 0.1
BEGIN

REGION Network 1: call generic code for the reject cylinder handler
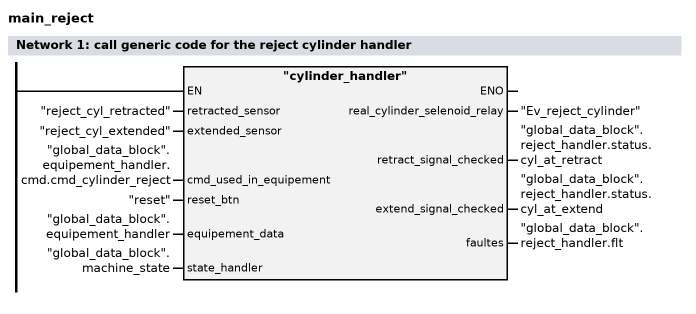
   RUNG wire#powerrail
      "cylinder_handler"(retracted_sensor := "reject_cyl_retracted", extended_sensor := "reject_cyl_extended", cmd_used_in_equipement := "global_data_block".equipement_handler.cmd.cmd_cylinder_reject, reset_btn := "reset", equipement_data := "global_data_block".equipement_handler, state_handler := "global_data_block".machine_state, real_cylinder_selenoid_relay => "Ev_reject_cylinder", retract_signal_checked => "global_data_block".reject_handler.status.cyl_at_retract, extend_signal_checked => "global_data_block".reject_handler.status.cyl_at_extend, faultes => "global_data_block".reject_handler.flt)
   END_RUNG
   // the same network as SCL:
   "cylinder_handler"(retracted_sensor := "reject_cyl_retracted",
                      extended_sensor := "reject_cyl_extended",
                      cmd_used_in_equipement := "global_data_block".equipement_handler.cmd.cmd_cylinder_reject,
                      reset_btn := "reset",
                      equipement_data := "global_data_block".equipement_handler,
                      state_handler := "global_data_block".machine_state,
                      real_cylinder_selenoid_relay => "Ev_reject_cylinder",
                      retract_signal_checked => "global_data_block".reject_handler.status.cyl_at_retract,
                      extend_signal_checked => "global_data_block".reject_handler.status.cyl_at_extend,
                      faultes => "global_data_block".reject_handler.flt);
END_REGION
END_FUNCTION

// folder: equipement/scaling

FUNCTION_BLOCK "scaling_sequence"   // FB10, LAD
{ S7_Optimized_Access := 'TRUE' }
VERSION : 0.1
   VAR_INPUT
      part_detect_scale : Bool;
      conveyer_feedbak : Bool;
   END_VAR
   VAR_IN_OUT
      equipement_handler : "udt_equipement";
      state_handler : "udt_state_handler";
      scaling_handler : "scaling_udt";
   END_VAR
   VAR
      start_conditon : Bool;
      state : Int;
      detected_bottle_weihgt : Int;
      weight_got : Bool;
      lock_verif_sequencer : Bool;
      IEC_Timer_0_Instance : TON_TIME;
   END_VAR
   VAR_TEMP
      verification_pulse : Bool;
      leaving_scale : Bool;
      part_detect_at_scale : Bool;
   END_VAR
   VAR_TEMP   // added for the SCL form of the ladder/FBD networks
      _w1 : Bool;
   END_VAR
BEGIN

REGION Network 1: define the start condition
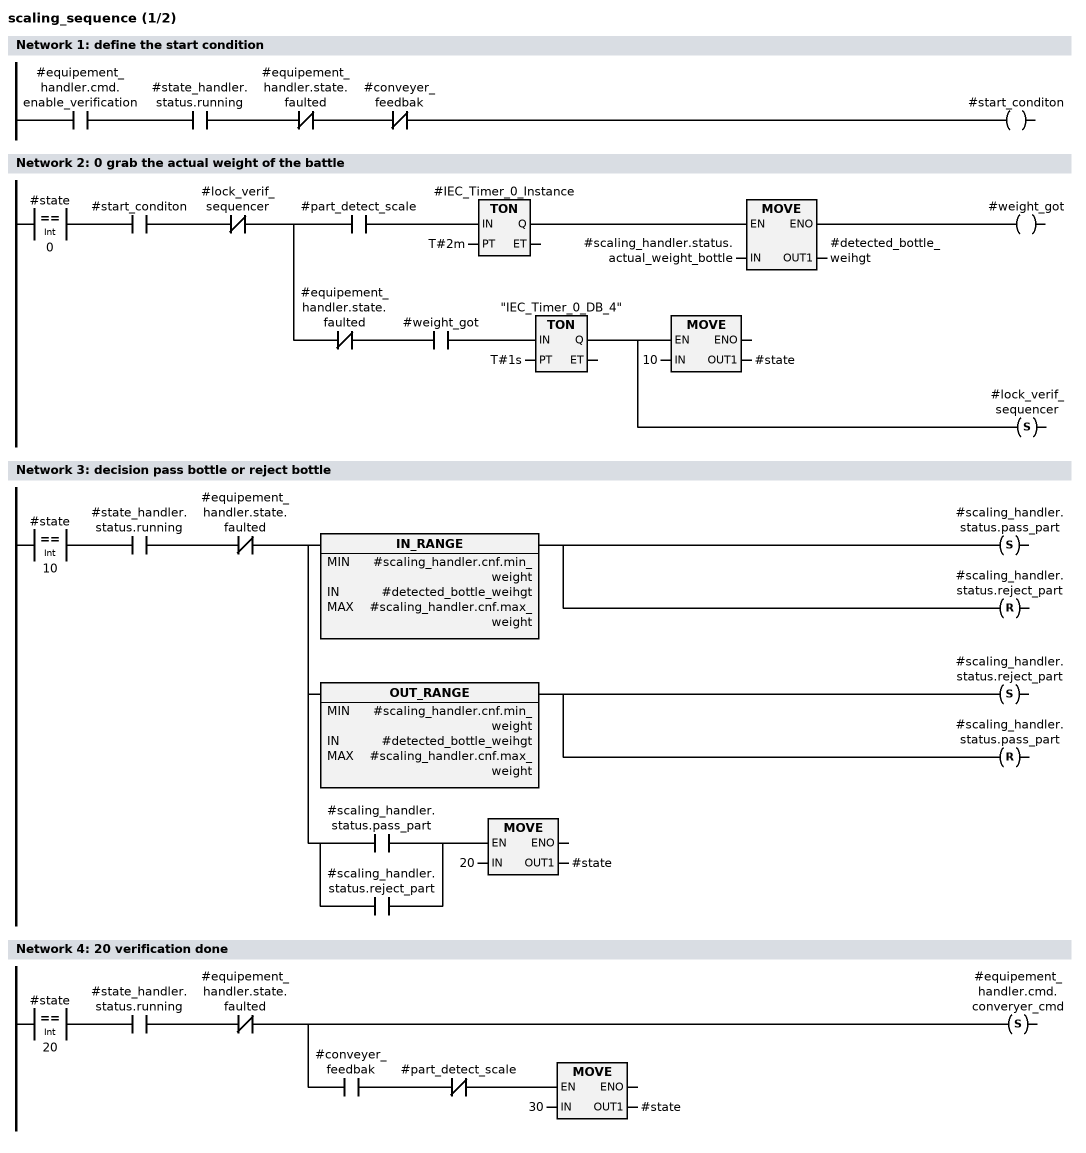
   RUNG wire#powerrail
      Contact( #equipement_handler.cmd.enable_verification )
      Contact( #state_handler.status.running )
      I_Contact( #equipement_handler.state.faulted )
      I_Contact( #conveyer_feedbak )
      Coil( #start_conditon )
   END_RUNG
   // the same network as SCL:
   #start_conditon := #equipement_handler.cmd.enable_verification AND #state_handler.status.running AND NOT #equipement_handler.state.faulted AND NOT #conveyer_feedbak;
END_REGION

REGION Network 2: 0 grab the actual weight of the battle
   #_w1 := (#state = 0) AND #start_conditon AND NOT #lock_verif_sequencer;
   #IEC_Timer_0_Instance(IN := #_w1 AND #part_detect_scale, PT := T#2m);   // TON
   IF #IEC_Timer_0_Instance.Q THEN
       #detected_bottle_weihgt := #scaling_handler.status.actual_weight_bottle;
   END_IF;
   #weight_got := #IEC_Timer_0_Instance.Q;
   "IEC_Timer_0_DB_4".TON(IN := #_w1 AND NOT #equipement_handler.state.faulted AND #weight_got, PT := T#1s);
   IF "IEC_Timer_0_DB_4".Q THEN
       #state := 10;
       #lock_verif_sequencer := TRUE;
   END_IF;
END_REGION

REGION Network 3: decision pass bottle or reject bottle
   #_w1 := (#state = 10) AND #state_handler.status.running AND NOT #equipement_handler.state.faulted;
   IF #_w1 AND (#scaling_handler.cnf.min_weight <= #detected_bottle_weihgt) AND (#detected_bottle_weihgt <= #scaling_handler.cnf.max_weight) THEN
       #scaling_handler.status.pass_part := TRUE;
       #scaling_handler.status.reject_part := FALSE;
   END_IF;
   IF #_w1 AND ((#detected_bottle_weihgt < #scaling_handler.cnf.min_weight) OR (#detected_bottle_weihgt > #scaling_handler.cnf.max_weight)) THEN
       #scaling_handler.status.reject_part := TRUE;
       #scaling_handler.status.pass_part := FALSE;
   END_IF;
   IF #_w1 AND (#scaling_handler.status.pass_part OR #scaling_handler.status.reject_part) THEN
       #state := 20;
   END_IF;
END_REGION

REGION Network 4: 20 verification done
   RUNG wire#powerrail
      { S7_Templates := "SrcType := Int" } EQ_Contact(in1 := #state, in2 := 20)
      Contact( #state_handler.status.running )
      I_Contact( #equipement_handler.state.faulted )
      wire#w1
      S_Coil( #equipement_handler.cmd.converyer_cmd )
   END_RUNG
   RUNG wire#w1
      Contact( #conveyer_feedbak )
      I_Contact( #part_detect_scale )
      Move(in := 30, out1 => #state)
   END_RUNG
   // the same network as SCL:
   #_w1 := (#state = 20) AND #state_handler.status.running AND NOT #equipement_handler.state.faulted;
   IF #_w1 THEN #equipement_handler.cmd.converyer_cmd := TRUE; END_IF;
   IF #_w1 AND #conveyer_feedbak AND NOT #part_detect_scale THEN #state := 30; END_IF;
END_REGION

REGION Network 5: 30 return to 0 and set the done_scaling check
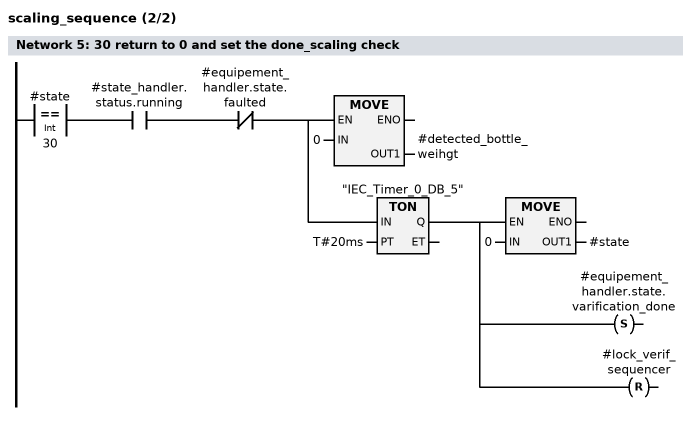
   #_w1 := (#state = 30) AND #state_handler.status.running AND NOT #equipement_handler.state.faulted;
   IF #_w1 THEN #detected_bottle_weihgt := 0; END_IF;
   "IEC_Timer_0_DB_5".TON(IN := #_w1, PT := T#20ms);
   IF "IEC_Timer_0_DB_5".Q THEN
       #state := 0;
       #equipement_handler.state.varification_done := TRUE;
       #lock_verif_sequencer := FALSE;
   END_IF;
END_REGION
END_FUNCTION_BLOCK

// folder: machine

FUNCTION_BLOCK "state_handler"   // FB2, LAD
{ S7_Optimized_Access := 'TRUE' }
VERSION : 0.1
// 0:ready
// 1:stop
// 2:running
// 3:faulted
   VAR_INPUT
      start_btn : Bool;
      reset_btn : Bool;
      stop_btn : Bool;
   END_VAR
   VAR_IN_OUT
      equipement_handler : "udt_equipement";
      state_handler : "udt_state_handler";
   END_VAR
   VAR_TEMP   // added for the SCL form of the ladder/FBD networks
      _w1 : Bool;
   END_VAR
BEGIN

REGION Network 1: transition from ready to running
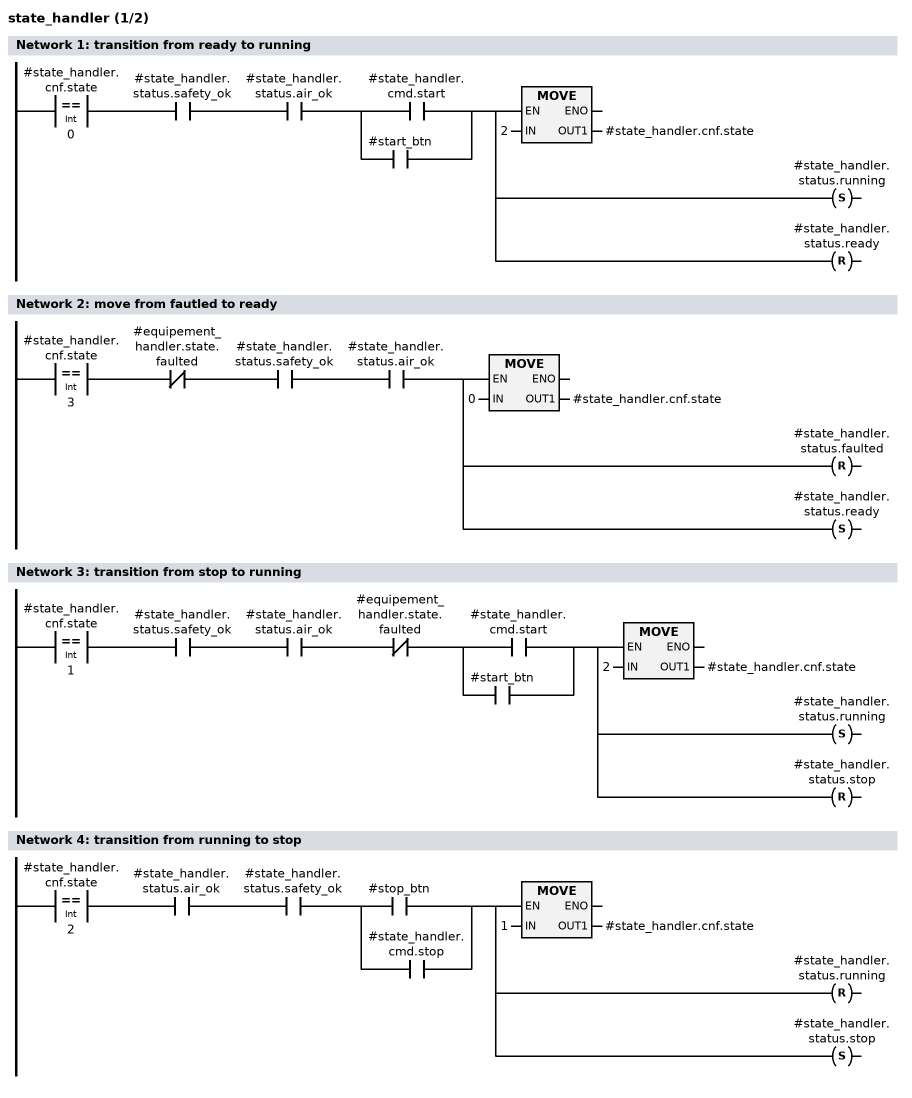
   RUNG wire#powerrail
      { S7_Templates := "SrcType := Int" } EQ_Contact(in1 := #state_handler.cnf.state, in2 := 0)
      Contact( #state_handler.status.safety_ok )
      Contact( #state_handler.status.air_ok )
      wire#w1
      Contact( #state_handler.cmd.start )
      wire#w2
      Move(in := 2, out1 => #state_handler.cnf.state)
   END_RUNG
   RUNG wire#w1
      Contact( #start_btn )
   END_RUNG wire#w2
   RUNG wire#w2
      S_Coil( #state_handler.status.running )
   END_RUNG
   RUNG wire#w2
      R_Coil( #state_handler.status.ready )
   END_RUNG
   // the same network as SCL:
   #_w1 := (#state_handler.cnf.state = 0) AND #state_handler.status.safety_ok AND #state_handler.status.air_ok AND (#state_handler.cmd.start OR #start_btn);
   IF #_w1 THEN
       #state_handler.cnf.state := 2;
       #state_handler.status.running := TRUE;
       #state_handler.status.ready := FALSE;
   END_IF;
END_REGION

REGION Network 2: move from fautled to ready
   RUNG wire#powerrail
      { S7_Templates := "SrcType := Int" } EQ_Contact(in1 := #state_handler.cnf.state, in2 := 3)
      I_Contact( #equipement_handler.state.faulted )
      Contact( #state_handler.status.safety_ok )
      Contact( #state_handler.status.air_ok )
      wire#w1
      Move(in := 0, out1 => #state_handler.cnf.state)
   END_RUNG
   RUNG wire#w1
      R_Coil( #state_handler.status.faulted )
   END_RUNG
   RUNG wire#w1
      S_Coil( #state_handler.status.ready )
   END_RUNG
   // the same network as SCL:
   #_w1 := (#state_handler.cnf.state = 3) AND NOT #equipement_handler.state.faulted AND #state_handler.status.safety_ok AND #state_handler.status.air_ok;
   IF #_w1 THEN
       #state_handler.cnf.state := 0;
       #state_handler.status.faulted := FALSE;
       #state_handler.status.ready := TRUE;
   END_IF;
END_REGION

REGION Network 3: transition from stop to running
   RUNG wire#powerrail
      { S7_Templates := "SrcType := Int" } EQ_Contact(in1 := #state_handler.cnf.state, in2 := 1)
      Contact( #state_handler.status.safety_ok )
      Contact( #state_handler.status.air_ok )
      I_Contact( #equipement_handler.state.faulted )
      wire#w1
      Contact( #state_handler.cmd.start )
      wire#w2
      Move(in := 2, out1 => #state_handler.cnf.state)
   END_RUNG
   RUNG wire#w1
      Contact( #start_btn )
   END_RUNG wire#w2
   RUNG wire#w2
      S_Coil( #state_handler.status.running )
   END_RUNG
   RUNG wire#w2
      R_Coil( #state_handler.status.stop )
   END_RUNG
   // the same network as SCL:
   #_w1 := (#state_handler.cnf.state = 1) AND #state_handler.status.safety_ok AND #state_handler.status.air_ok AND NOT #equipement_handler.state.faulted AND (#state_handler.cmd.start OR #start_btn);
   IF #_w1 THEN
       #state_handler.cnf.state := 2;
       #state_handler.status.running := TRUE;
       #state_handler.status.stop := FALSE;
   END_IF;
END_REGION

REGION Network 4: transition from running to stop
   RUNG wire#powerrail
      { S7_Templates := "SrcType := Int" } EQ_Contact(in1 := #state_handler.cnf.state, in2 := 2)
      Contact( #state_handler.status.air_ok )
      Contact( #state_handler.status.safety_ok )
      wire#w1
      Contact( #stop_btn )
      wire#w2
      Move(in := 1, out1 => #state_handler.cnf.state)
   END_RUNG
   RUNG wire#w1
      Contact( #state_handler.cmd.stop )
   END_RUNG wire#w2
   RUNG wire#w2
      R_Coil( #state_handler.status.running )
   END_RUNG
   RUNG wire#w2
      S_Coil( #state_handler.status.stop )
   END_RUNG
   // the same network as SCL:
   #_w1 := (#state_handler.cnf.state = 2) AND #state_handler.status.air_ok AND #state_handler.status.safety_ok AND (#stop_btn OR #state_handler.cmd.stop);
   IF #_w1 THEN
       #state_handler.cnf.state := 1;
       #state_handler.status.running := FALSE;
       #state_handler.status.stop := TRUE;
   END_IF;
END_REGION

REGION Network 5: transition from any state to faulted
